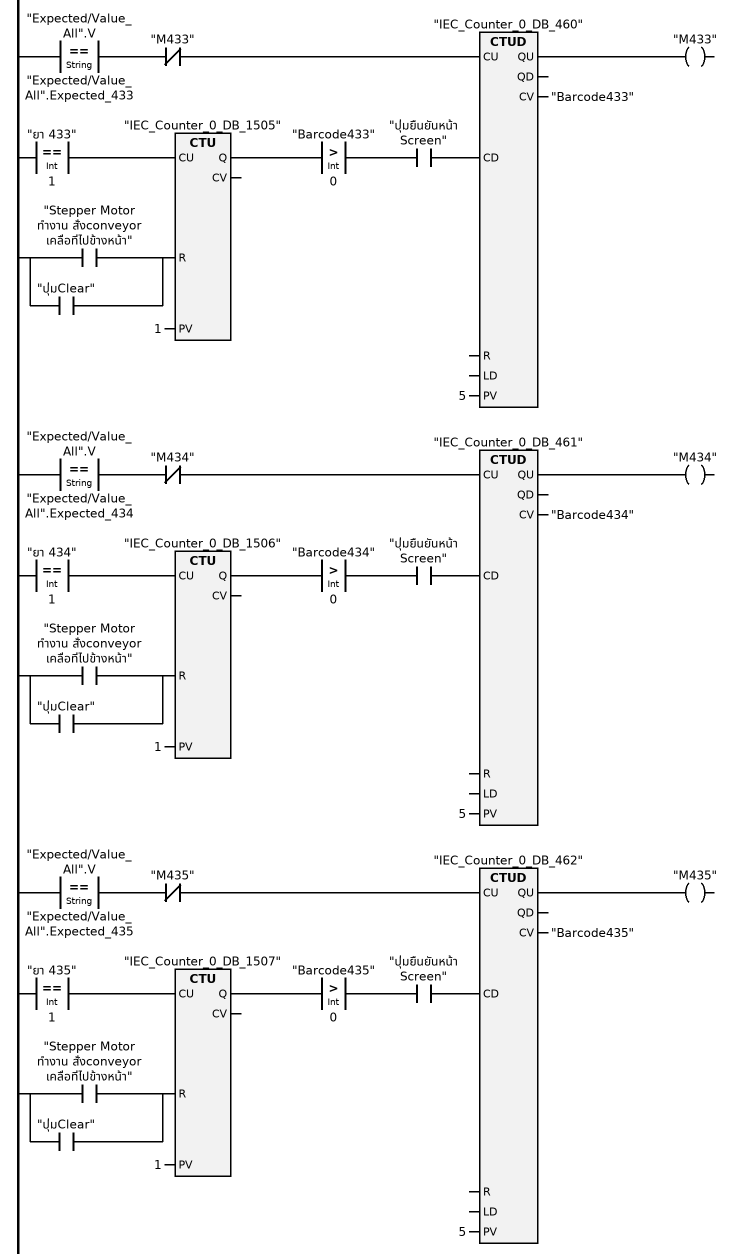
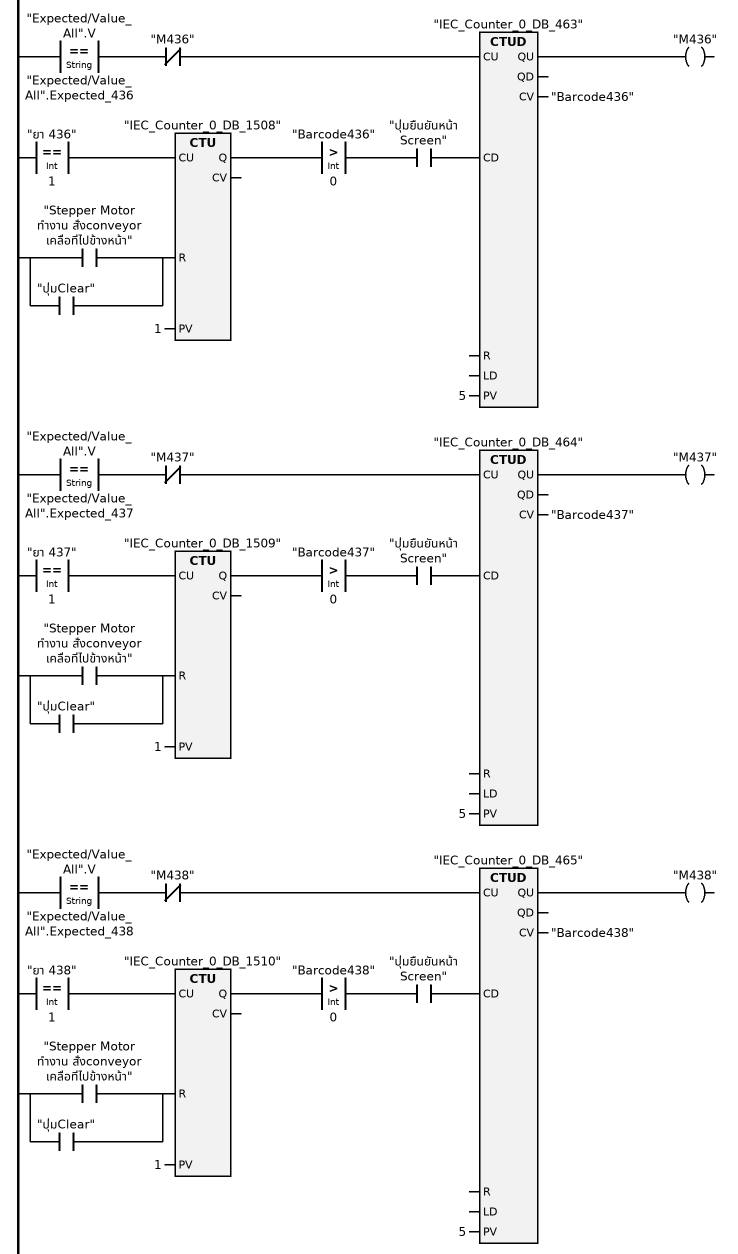
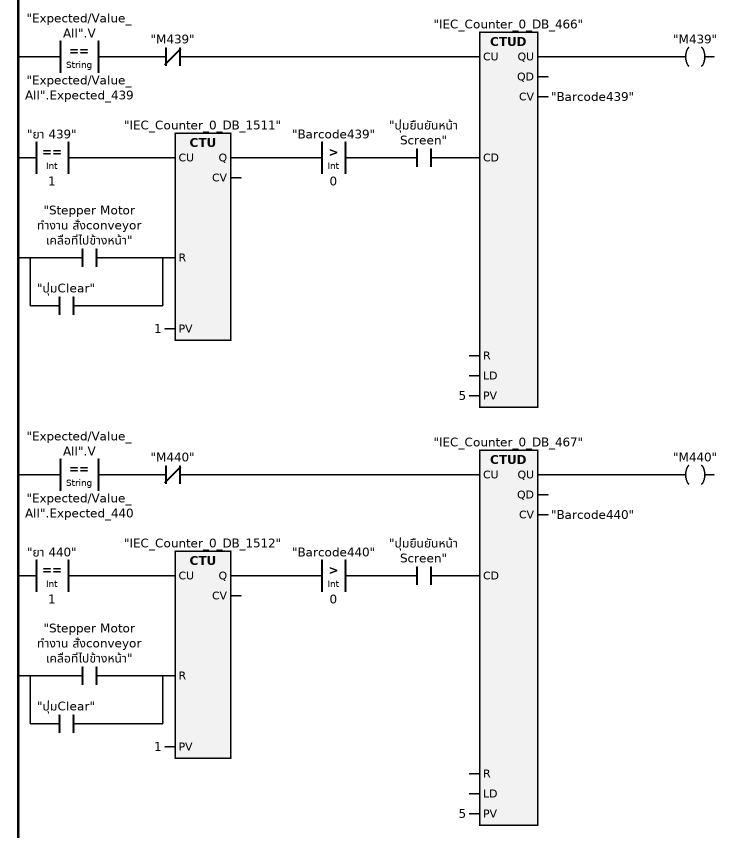
   "IEC_Counter_0_DB_1493".CTU(CU := "ยา 421" = 1,
                           R := "Stepper Motor ทำงาน สั่งconveyor เคลื่อที่ไปข้างหน้า" OR "ปุ่มClear",
                           PV := 1);
   "IEC_Counter_0_DB_448".CTUD(CU := ("Expected/Value_All".V = "Expected/Value_All".Expected_421) AND NOT "M421",
                           CD := "IEC_Counter_0_DB_1493".Q AND ("Barcode421" > 0) AND "ปุ่มยืนยันหน้า Screen",
                           PV := 5,
                           CV => "Barcode421");
   "M421" := "IEC_Counter_0_DB_448".QU;
   "IEC_Counter_0_DB_1494".CTU(CU := "ยา 422" = 1,
                           R := "Stepper Motor ทำงาน สั่งconveyor เคลื่อที่ไปข้างหน้า" OR "ปุ่มClear",
                           PV := 1);
   "IEC_Counter_0_DB_449".CTUD(CU := ("Expected/Value_All".V = "Expected/Value_All".Expected_422) AND NOT "M422",
                           CD := "IEC_Counter_0_DB_1494".Q AND ("Barcode422" > 0) AND "ปุ่มยืนยันหน้า Screen",
                           PV := 5,
                           CV => "Barcode422");
   "M422" := "IEC_Counter_0_DB_449".QU;
   "IEC_Counter_0_DB_1495".CTU(CU := "ยา 423" = 1,
                           R := "Stepper Motor ทำงาน สั่งconveyor เคลื่อที่ไปข้างหน้า" OR "ปุ่มClear",
                           PV := 1);
   "IEC_Counter_0_DB_450".CTUD(CU := ("Expected/Value_All".V = "Expected/Value_All".Expected_423) AND NOT "M423",
                           CD := "IEC_Counter_0_DB_1495".Q AND ("Barcode423" > 0) AND "ปุ่มยืนยันหน้า Screen",
                           PV := 5,
                           CV => "Barcode423");
   "M423" := "IEC_Counter_0_DB_450".QU;
   "IEC_Counter_0_DB_1496".CTU(CU := "ยา 424" = 1,
                           R := "Stepper Motor ทำงาน สั่งconveyor เคลื่อที่ไปข้างหน้า" OR "ปุ่มClear",
                           PV := 1);
   "IEC_Counter_0_DB_451".CTUD(CU := ("Expected/Value_All".V = "Expected/Value_All".Expected_424) AND NOT "M424",
                           CD := "IEC_Counter_0_DB_1496".Q AND ("Barcode424" > 0) AND "ปุ่มยืนยันหน้า Screen",
                           PV := 5,
                           CV => "Barcode424");
   "M424" := "IEC_Counter_0_DB_451".QU;
   "IEC_Counter_0_DB_1497".CTU(CU := "ยา 425" = 1,
                           R := "Stepper Motor ทำงาน สั่งconveyor เคลื่อที่ไปข้างหน้า" OR "ปุ่มClear",
                           PV := 1);
   "IEC_Counter_0_DB_452".CTUD(CU := ("Expected/Value_All".V = "Expected/Value_All".Expected_425) AND NOT "M425",
                           CD := "IEC_Counter_0_DB_1497".Q AND ("Barcode425" > 0) AND "ปุ่มยืนยันหน้า Screen",
                           PV := 5,
                           CV => "Barcode425");
   "M425" := "IEC_Counter_0_DB_452".QU;
   "IEC_Counter_0_DB_1498".CTU(CU := "ยา 426" = 1,
                           R := "Stepper Motor ทำงาน สั่งconveyor เคลื่อที่ไปข้างหน้า" OR "ปุ่มClear",
                           PV := 1);
   "IEC_Counter_0_DB_453".CTUD(CU := ("Expected/Value_All".V = "Expected/Value_All".Expected_426) AND NOT "M426",
                           CD := "IEC_Counter_0_DB_1498".Q AND ("Barcode426" > 0) AND "ปุ่มยืนยันหน้า Screen",
                           PV := 5,
                           CV => "Barcode426");
   "M426" := "IEC_Counter_0_DB_453".QU;
   "IEC_Counter_0_DB_1499".CTU(CU := "ยา 427" = 1,
                           R := "Stepper Motor ทำงาน สั่งconveyor เคลื่อที่ไปข้างหน้า" OR "ปุ่มClear",
                           PV := 1);
   "IEC_Counter_0_DB_454".CTUD(CU := ("Expected/Value_All".V = "Expected/Value_All".Expected_427) AND NOT "M427",
                           CD := "IEC_Counter_0_DB_1499".Q AND ("Barcode427" > 0) AND "ปุ่มยืนยันหน้า Screen",
                           PV := 5,
                           CV => "Barcode427");
   "M427" := "IEC_Counter_0_DB_454".QU;
   "IEC_Counter_0_DB_1500".CTU(CU := "ยา 428" = 1,
                           R := "Stepper Motor ทำงาน สั่งconveyor เคลื่อที่ไปข้างหน้า" OR "ปุ่มClear",
                           PV := 1);
   "IEC_Counter_0_DB_455".CTUD(CU := ("Expected/Value_All".V = "Expected/Value_All".Expected_428) AND NOT "M428",
                           CD := "IEC_Counter_0_DB_1500".Q AND ("Barcode428" > 0) AND "ปุ่มยืนยันหน้า Screen",
                           PV := 5,
                           CV => "Barcode428");
   "M428" := "IEC_Counter_0_DB_455".QU;
   "IEC_Counter_0_DB_1501".CTU(CU := "ยา 429" = 1,
                           R := "Stepper Motor ทำงาน สั่งconveyor เคลื่อที่ไปข้างหน้า" OR "ปุ่มClear",
                           PV := 1);
   "IEC_Counter_0_DB_456".CTUD(CU := ("Expected/Value_All".V = "Expected/Value_All".Expected_429) AND NOT "M429",
                           CD := "IEC_Counter_0_DB_1501".Q AND ("Barcode429" > 0) AND "ปุ่มยืนยันหน้า Screen",
                           PV := 5,
                           CV => "Barcode429");
   "M429" := "IEC_Counter_0_DB_456".QU;
   "IEC_Counter_0_DB_1502".CTU(CU := "ยา 430" = 1,
                           R := "Stepper Motor ทำงาน สั่งconveyor เคลื่อที่ไปข้างหน้า" OR "ปุ่มClear",
                           PV := 1);
   "IEC_Counter_0_DB_457".CTUD(CU := ("Expected/Value_All".V = "Expected/Value_All".Expected_430) AND NOT "M430",
                           CD := "IEC_Counter_0_DB_1502".Q AND ("Barcode430" > 0) AND "ปุ่มยืนยันหน้า Screen",
                           PV := 5,
                           CV => "Barcode430");
   "M430" := "IEC_Counter_0_DB_457".QU;
   "IEC_Counter_0_DB_1503".CTU(CU := "ยา 431" = 1,
                           R := "Stepper Motor ทำงาน สั่งconveyor เคลื่อที่ไปข้างหน้า" OR "ปุ่มClear",
                           PV := 1);
   "IEC_Counter_0_DB_458".CTUD(CU := ("Expected/Value_All".V = "Expected/Value_All".Expected_431) AND NOT "M431",
                           CD := "IEC_Counter_0_DB_1503".Q AND ("Barcode431" > 0) AND "ปุ่มยืนยันหน้า Screen",
                           PV := 5,
                           CV => "Barcode431");
   "M431" := "IEC_Counter_0_DB_458".QU;
   "IEC_Counter_0_DB_1504".CTU(CU := "ยา 432" = 1,
                           R := "Stepper Motor ทำงาน สั่งconveyor เคลื่อที่ไปข้างหน้า" OR "ปุ่มClear",
                           PV := 1);
   "IEC_Counter_0_DB_459".CTUD(CU := ("Expected/Value_All".V = "Expected/Value_All".Expected_432) AND NOT "M432",
                           CD := "IEC_Counter_0_DB_1504".Q AND ("Barcode432" > 0) AND "ปุ่มยืนยันหน้า Screen",
                           PV := 5,
                           CV => "Barcode432");
   "M432" := "IEC_Counter_0_DB_459".QU;
   "IEC_Counter_0_DB_1505".CTU(CU := "ยา 433" = 1,
                           R := "Stepper Motor ทำงาน สั่งconveyor เคลื่อที่ไปข้างหน้า" OR "ปุ่มClear",
                           PV := 1);
   "IEC_Counter_0_DB_460".CTUD(CU := ("Expected/Value_All".V = "Expected/Value_All".Expected_433) AND NOT "M433",
                           CD := "IEC_Counter_0_DB_1505".Q AND ("Barcode433" > 0) AND "ปุ่มยืนยันหน้า Screen",
                           PV := 5,
                           CV => "Barcode433");
   "M433" := "IEC_Counter_0_DB_460".QU;
   "IEC_Counter_0_DB_1506".CTU(CU := "ยา 434" = 1,
                           R := "Stepper Motor ทำงาน สั่งconveyor เคลื่อที่ไปข้างหน้า" OR "ปุ่มClear",
                           PV := 1);
   "IEC_Counter_0_DB_461".CTUD(CU := ("Expected/Value_All".V = "Expected/Value_All".Expected_434) AND NOT "M434",
                           CD := "IEC_Counter_0_DB_1506".Q AND ("Barcode434" > 0) AND "ปุ่มยืนยันหน้า Screen",
                           PV := 5,
                           CV => "Barcode434");
   "M434" := "IEC_Counter_0_DB_461".QU;
   "IEC_Counter_0_DB_1507".CTU(CU := "ยา 435" = 1,
                           R := "Stepper Motor ทำงาน สั่งconveyor เคลื่อที่ไปข้างหน้า" OR "ปุ่มClear",
                           PV := 1);
   "IEC_Counter_0_DB_462".CTUD(CU := ("Expected/Value_All".V = "Expected/Value_All".Expected_435) AND NOT "M435",
                           CD := "IEC_Counter_0_DB_1507".Q AND ("Barcode435" > 0) AND "ปุ่มยืนยันหน้า Screen",
                           PV := 5,
                           CV => "Barcode435");
   "M435" := "IEC_Counter_0_DB_462".QU;
   "IEC_Counter_0_DB_1508".CTU(CU := "ยา 436" = 1,
                           R := "Stepper Motor ทำงาน สั่งconveyor เคลื่อที่ไปข้างหน้า" OR "ปุ่มClear",
                           PV := 1);
   "IEC_Counter_0_DB_463".CTUD(CU := ("Expected/Value_All".V = "Expected/Value_All".Expected_436) AND NOT "M436",
                           CD := "IEC_Counter_0_DB_1508".Q AND ("Barcode436" > 0) AND "ปุ่มยืนยันหน้า Screen",
                           PV := 5,
                           CV => "Barcode436");
   "M436" := "IEC_Counter_0_DB_463".QU;
   "IEC_Counter_0_DB_1509".CTU(CU := "ยา 437" = 1,
                           R := "Stepper Motor ทำงาน สั่งconveyor เคลื่อที่ไปข้างหน้า" OR "ปุ่มClear",
                           PV := 1);
   "IEC_Counter_0_DB_464".CTUD(CU := ("Expected/Value_All".V = "Expected/Value_All".Expected_437) AND NOT "M437",
                           CD := "IEC_Counter_0_DB_1509".Q AND ("Barcode437" > 0) AND "ปุ่มยืนยันหน้า Screen",
                           PV := 5,
                           CV => "Barcode437");
   "M437" := "IEC_Counter_0_DB_464".QU;
   "IEC_Counter_0_DB_1510".CTU(CU := "ยา 438" = 1,
                           R := "Stepper Motor ทำงาน สั่งconveyor เคลื่อที่ไปข้างหน้า" OR "ปุ่มClear",
                           PV := 1);
   "IEC_Counter_0_DB_465".CTUD(CU := ("Expected/Value_All".V = "Expected/Value_All".Expected_438) AND NOT "M438",
                           CD := "IEC_Counter_0_DB_1510".Q AND ("Barcode438" > 0) AND "ปุ่มยืนยันหน้า Screen",
                           PV := 5,
                           CV => "Barcode438");
   "M438" := "IEC_Counter_0_DB_465".QU;
   "IEC_Counter_0_DB_1511".CTU(CU := "ยา 439" = 1,
                           R := "Stepper Motor ทำงาน สั่งconveyor เคลื่อที่ไปข้างหน้า" OR "ปุ่มClear",
                           PV := 1);
   "IEC_Counter_0_DB_466".CTUD(CU := ("Expected/Value_All".V = "Expected/Value_All".Expected_439) AND NOT "M439",
                           CD := "IEC_Counter_0_DB_1511".Q AND ("Barcode439" > 0) AND "ปุ่มยืนยันหน้า Screen",
                           PV := 5,
                           CV => "Barcode439");
   "M439" := "IEC_Counter_0_DB_466".QU;
   "IEC_Counter_0_DB_1512".CTU(CU := "ยา 440" = 1,
                           R := "Stepper Motor ทำงาน สั่งconveyor เคลื่อที่ไปข้างหน้า" OR "ปุ่มClear",
                           PV := 1);
   "IEC_Counter_0_DB_467".CTUD(CU := ("Expected/Value_All".V = "Expected/Value_All".Expected_440) AND NOT "M440",
                           CD := "IEC_Counter_0_DB_1512".Q AND ("Barcode440" > 0) AND "ปุ่มยืนยันหน้า Screen",
                           PV := 5,
                           CV => "Barcode440");
   "M440" := "IEC_Counter_0_DB_467".QU;
END_REGION

REGION Network 23
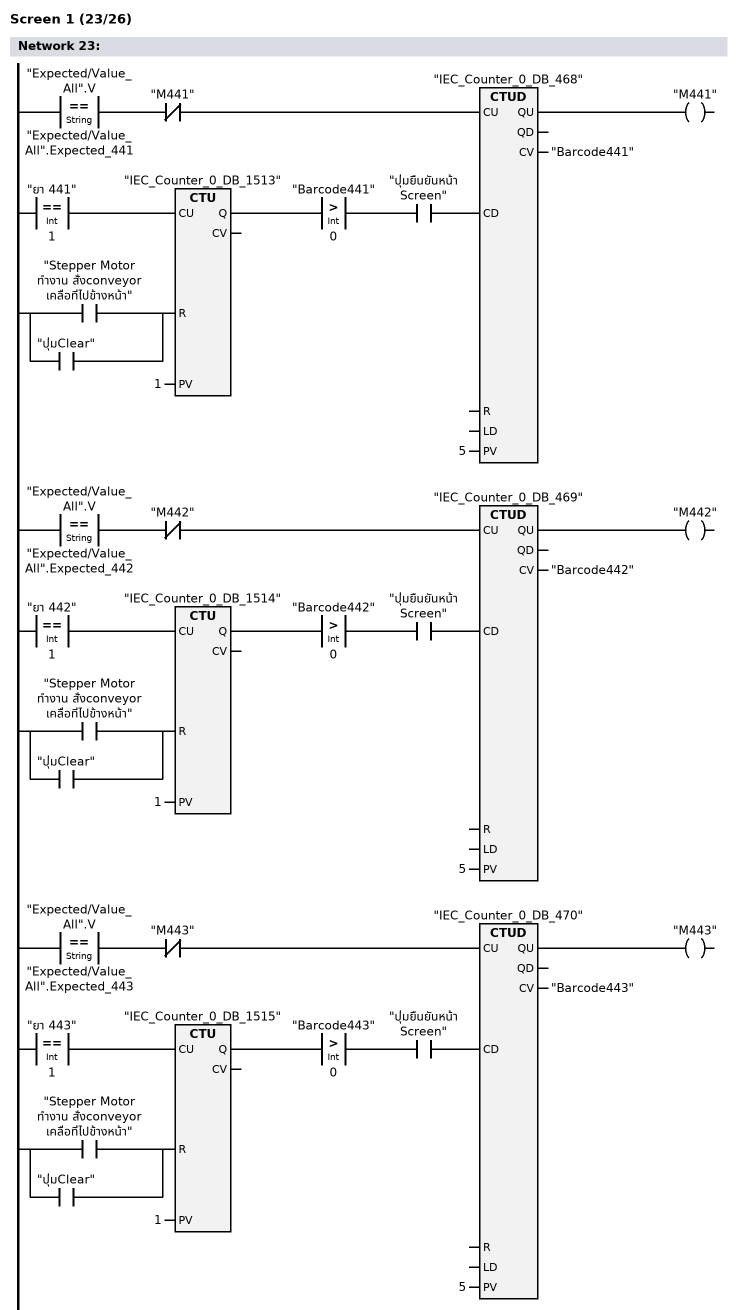
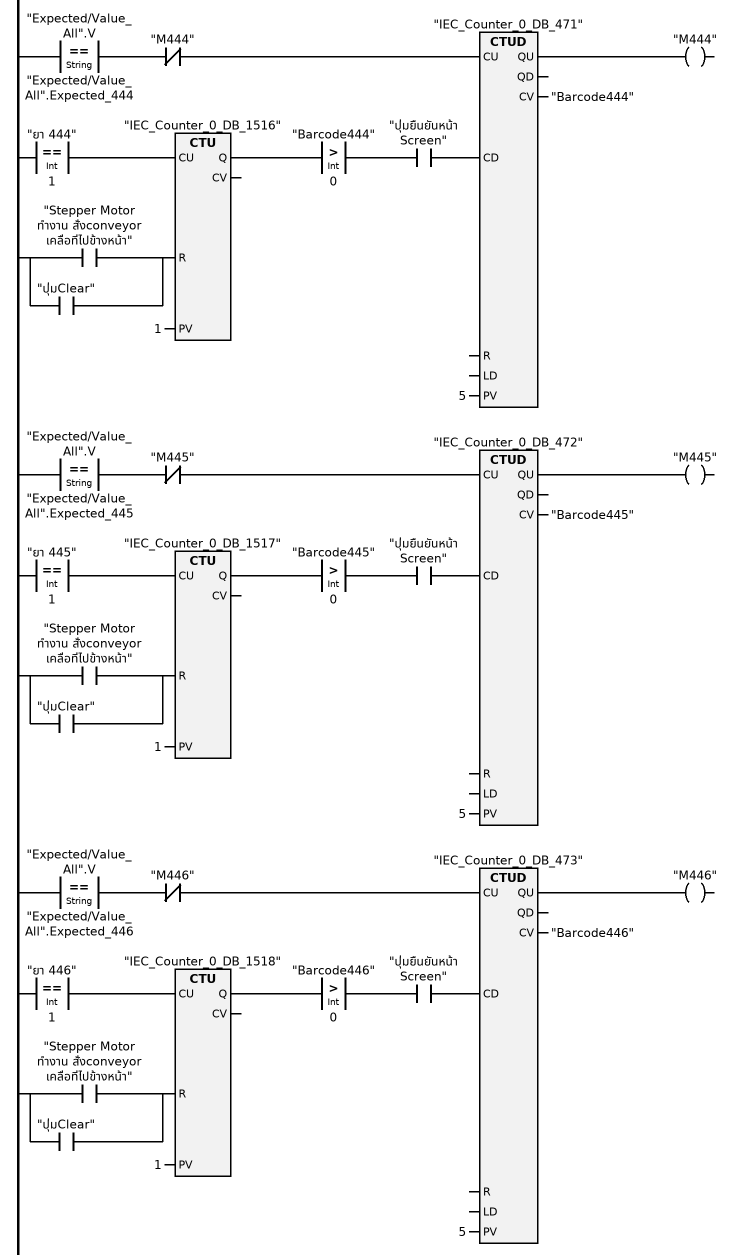
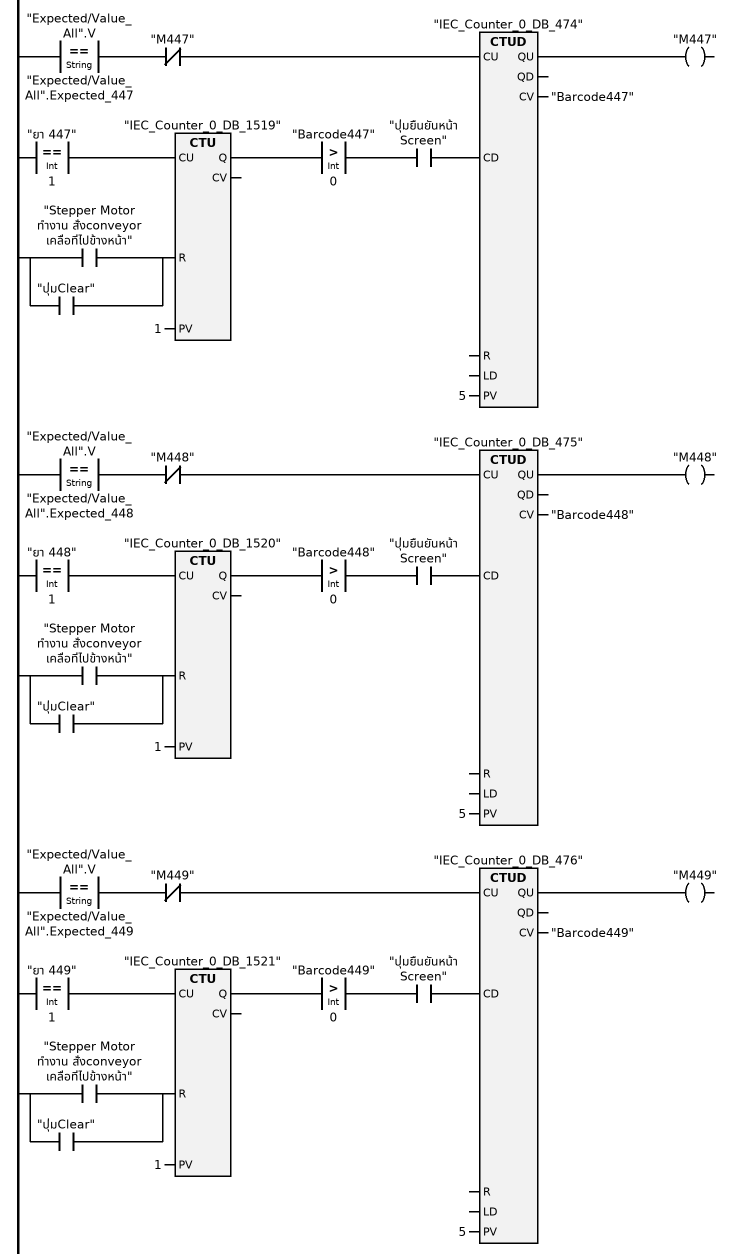
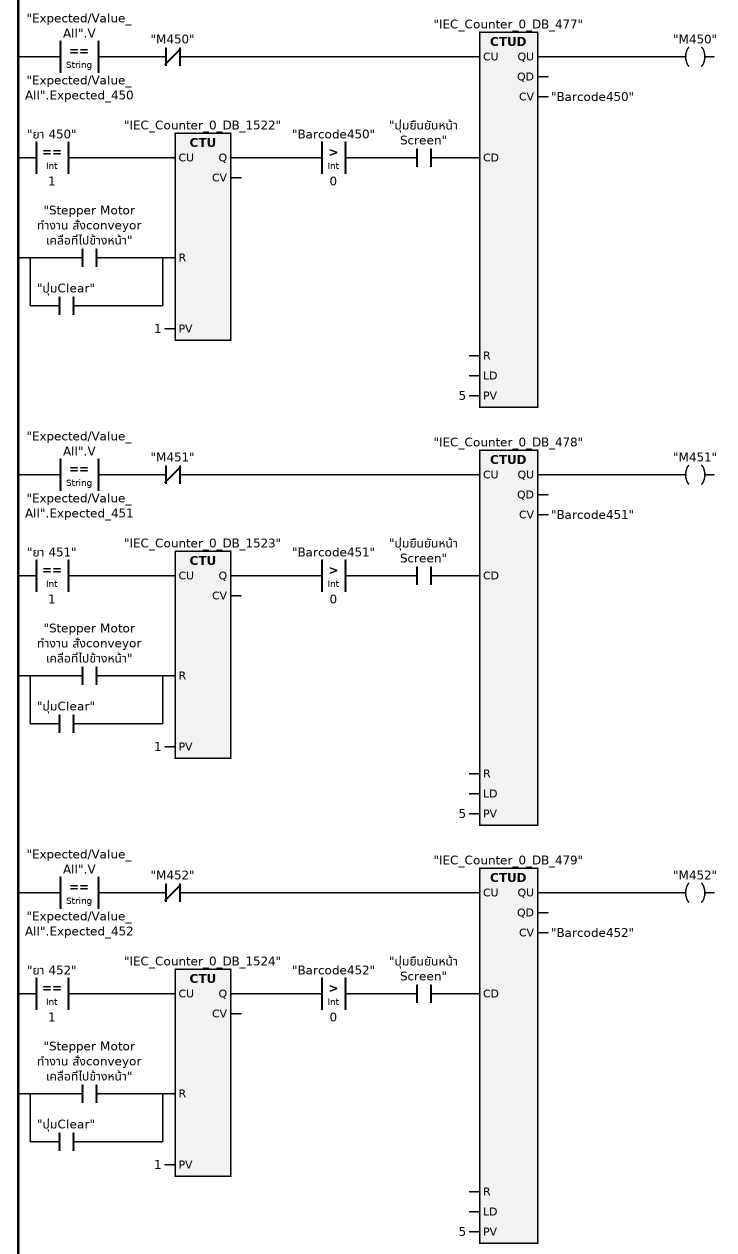
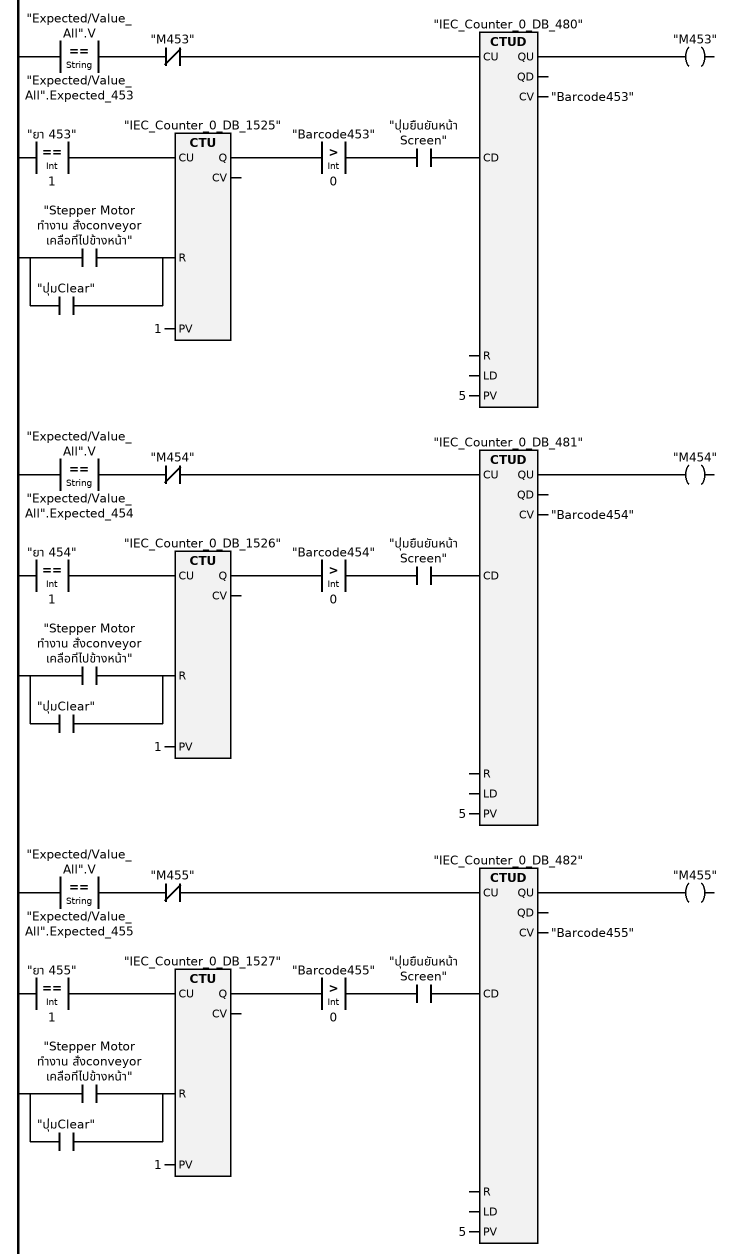
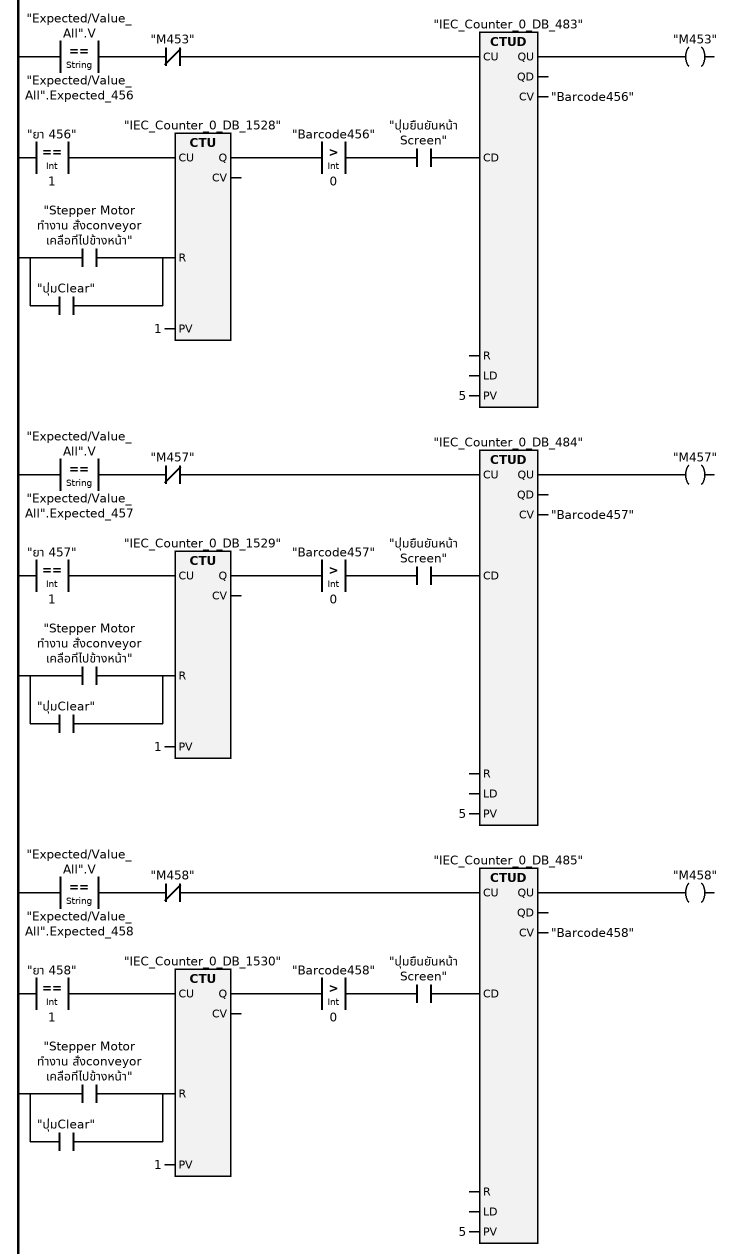
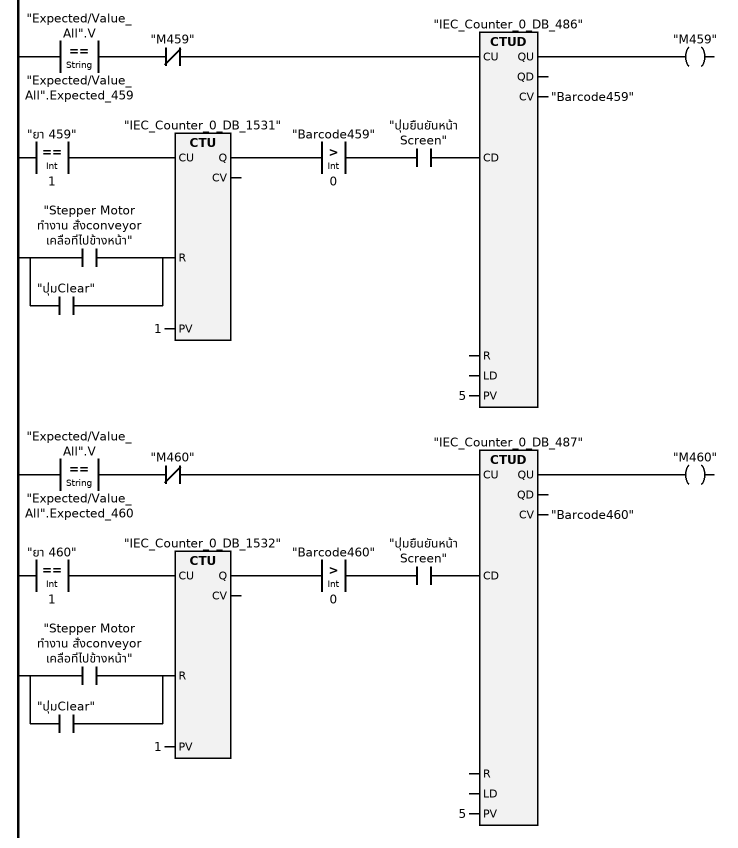
   "IEC_Counter_0_DB_1513".CTU(CU := "ยา 441" = 1,
                           R := "Stepper Motor ทำงาน สั่งconveyor เคลื่อที่ไปข้างหน้า" OR "ปุ่มClear",
                           PV := 1);
   "IEC_Counter_0_DB_468".CTUD(CU := ("Expected/Value_All".V = "Expected/Value_All".Expected_441) AND NOT "M441",
                           CD := "IEC_Counter_0_DB_1513".Q AND ("Barcode441" > 0) AND "ปุ่มยืนยันหน้า Screen",
                           PV := 5,
                           CV => "Barcode441");
   "M441" := "IEC_Counter_0_DB_468".QU;
   "IEC_Counter_0_DB_1514".CTU(CU := "ยา 442" = 1,
                           R := "Stepper Motor ทำงาน สั่งconveyor เคลื่อที่ไปข้างหน้า" OR "ปุ่มClear",
                           PV := 1);
   "IEC_Counter_0_DB_469".CTUD(CU := ("Expected/Value_All".V = "Expected/Value_All".Expected_442) AND NOT "M442",
                           CD := "IEC_Counter_0_DB_1514".Q AND ("Barcode442" > 0) AND "ปุ่มยืนยันหน้า Screen",
                           PV := 5,
                           CV => "Barcode442");
   "M442" := "IEC_Counter_0_DB_469".QU;
   "IEC_Counter_0_DB_1515".CTU(CU := "ยา 443" = 1,
                           R := "Stepper Motor ทำงาน สั่งconveyor เคลื่อที่ไปข้างหน้า" OR "ปุ่มClear",
                           PV := 1);
   "IEC_Counter_0_DB_470".CTUD(CU := ("Expected/Value_All".V = "Expected/Value_All".Expected_443) AND NOT "M443",
                           CD := "IEC_Counter_0_DB_1515".Q AND ("Barcode443" > 0) AND "ปุ่มยืนยันหน้า Screen",
                           PV := 5,
                           CV => "Barcode443");
   "M443" := "IEC_Counter_0_DB_470".QU;
   "IEC_Counter_0_DB_1516".CTU(CU := "ยา 444" = 1,
                           R := "Stepper Motor ทำงาน สั่งconveyor เคลื่อที่ไปข้างหน้า" OR "ปุ่มClear",
                           PV := 1);
   "IEC_Counter_0_DB_471".CTUD(CU := ("Expected/Value_All".V = "Expected/Value_All".Expected_444) AND NOT "M444",
                           CD := "IEC_Counter_0_DB_1516".Q AND ("Barcode444" > 0) AND "ปุ่มยืนยันหน้า Screen",
                           PV := 5,
                           CV => "Barcode444");
   "M444" := "IEC_Counter_0_DB_471".QU;
   "IEC_Counter_0_DB_1517".CTU(CU := "ยา 445" = 1,
                           R := "Stepper Motor ทำงาน สั่งconveyor เคลื่อที่ไปข้างหน้า" OR "ปุ่มClear",
                           PV := 1);
   "IEC_Counter_0_DB_472".CTUD(CU := ("Expected/Value_All".V = "Expected/Value_All".Expected_445) AND NOT "M445",
                           CD := "IEC_Counter_0_DB_1517".Q AND ("Barcode445" > 0) AND "ปุ่มยืนยันหน้า Screen",
                           PV := 5,
                           CV => "Barcode445");
   "M445" := "IEC_Counter_0_DB_472".QU;
   "IEC_Counter_0_DB_1518".CTU(CU := "ยา 446" = 1,
                           R := "Stepper Motor ทำงาน สั่งconveyor เคลื่อที่ไปข้างหน้า" OR "ปุ่มClear",
                           PV := 1);
   "IEC_Counter_0_DB_473".CTUD(CU := ("Expected/Value_All".V = "Expected/Value_All".Expected_446) AND NOT "M446",
                           CD := "IEC_Counter_0_DB_1518".Q AND ("Barcode446" > 0) AND "ปุ่มยืนยันหน้า Screen",
                           PV := 5,
                           CV => "Barcode446");
   "M446" := "IEC_Counter_0_DB_473".QU;
   "IEC_Counter_0_DB_1519".CTU(CU := "ยา 447" = 1,
                           R := "Stepper Motor ทำงาน สั่งconveyor เคลื่อที่ไปข้างหน้า" OR "ปุ่มClear",
                           PV := 1);
   "IEC_Counter_0_DB_474".CTUD(CU := ("Expected/Value_All".V = "Expected/Value_All".Expected_447) AND NOT "M447",
                           CD := "IEC_Counter_0_DB_1519".Q AND ("Barcode447" > 0) AND "ปุ่มยืนยันหน้า Screen",
                           PV := 5,
                           CV => "Barcode447");
   "M447" := "IEC_Counter_0_DB_474".QU;
   "IEC_Counter_0_DB_1520".CTU(CU := "ยา 448" = 1,
                           R := "Stepper Motor ทำงาน สั่งconveyor เคลื่อที่ไปข้างหน้า" OR "ปุ่มClear",
                           PV := 1);
   "IEC_Counter_0_DB_475".CTUD(CU := ("Expected/Value_All".V = "Expected/Value_All".Expected_448) AND NOT "M448",
                           CD := "IEC_Counter_0_DB_1520".Q AND ("Barcode448" > 0) AND "ปุ่มยืนยันหน้า Screen",
                           PV := 5,
                           CV => "Barcode448");
   "M448" := "IEC_Counter_0_DB_475".QU;
   "IEC_Counter_0_DB_1521".CTU(CU := "ยา 449" = 1,
                           R := "Stepper Motor ทำงาน สั่งconveyor เคลื่อที่ไปข้างหน้า" OR "ปุ่มClear",
                           PV := 1);
   "IEC_Counter_0_DB_476".CTUD(CU := ("Expected/Value_All".V = "Expected/Value_All".Expected_449) AND NOT "M449",
                           CD := "IEC_Counter_0_DB_1521".Q AND ("Barcode449" > 0) AND "ปุ่มยืนยันหน้า Screen",
                           PV := 5,
                           CV => "Barcode449");
   "M449" := "IEC_Counter_0_DB_476".QU;
   "IEC_Counter_0_DB_1522".CTU(CU := "ยา 450" = 1,
                           R := "Stepper Motor ทำงาน สั่งconveyor เคลื่อที่ไปข้างหน้า" OR "ปุ่มClear",
                           PV := 1);
   "IEC_Counter_0_DB_477".CTUD(CU := ("Expected/Value_All".V = "Expected/Value_All".Expected_450) AND NOT "M450",
                           CD := "IEC_Counter_0_DB_1522".Q AND ("Barcode450" > 0) AND "ปุ่มยืนยันหน้า Screen",
                           PV := 5,
                           CV => "Barcode450");
   "M450" := "IEC_Counter_0_DB_477".QU;
   "IEC_Counter_0_DB_1523".CTU(CU := "ยา 451" = 1,
                           R := "Stepper Motor ทำงาน สั่งconveyor เคลื่อที่ไปข้างหน้า" OR "ปุ่มClear",
                           PV := 1);
   "IEC_Counter_0_DB_478".CTUD(CU := ("Expected/Value_All".V = "Expected/Value_All".Expected_451) AND NOT "M451",
                           CD := "IEC_Counter_0_DB_1523".Q AND ("Barcode451" > 0) AND "ปุ่มยืนยันหน้า Screen",
                           PV := 5,
                           CV => "Barcode451");
   "M451" := "IEC_Counter_0_DB_478".QU;
   "IEC_Counter_0_DB_1524".CTU(CU := "ยา 452" = 1,
                           R := "Stepper Motor ทำงาน สั่งconveyor เคลื่อที่ไปข้างหน้า" OR "ปุ่มClear",
                           PV := 1);
   "IEC_Counter_0_DB_479".CTUD(CU := ("Expected/Value_All".V = "Expected/Value_All".Expected_452) AND NOT "M452",
                           CD := "IEC_Counter_0_DB_1524".Q AND ("Barcode452" > 0) AND "ปุ่มยืนยันหน้า Screen",
                           PV := 5,
                           CV => "Barcode452");
   "M452" := "IEC_Counter_0_DB_479".QU;
   "IEC_Counter_0_DB_1525".CTU(CU := "ยา 453" = 1,
                           R := "Stepper Motor ทำงาน สั่งconveyor เคลื่อที่ไปข้างหน้า" OR "ปุ่มClear",
                           PV := 1);
   "IEC_Counter_0_DB_480".CTUD(CU := ("Expected/Value_All".V = "Expected/Value_All".Expected_453) AND NOT "M453",
                           CD := "IEC_Counter_0_DB_1525".Q AND ("Barcode453" > 0) AND "ปุ่มยืนยันหน้า Screen",
                           PV := 5,
                           CV => "Barcode453");
   "M453" := "IEC_Counter_0_DB_480".QU;
   "IEC_Counter_0_DB_1526".CTU(CU := "ยา 454" = 1,
                           R := "Stepper Motor ทำงาน สั่งconveyor เคลื่อที่ไปข้างหน้า" OR "ปุ่มClear",
                           PV := 1);
   "IEC_Counter_0_DB_481".CTUD(CU := ("Expected/Value_All".V = "Expected/Value_All".Expected_454) AND NOT "M454",
                           CD := "IEC_Counter_0_DB_1526".Q AND ("Barcode454" > 0) AND "ปุ่มยืนยันหน้า Screen",
                           PV := 5,
                           CV => "Barcode454");
   "M454" := "IEC_Counter_0_DB_481".QU;
   "IEC_Counter_0_DB_1527".CTU(CU := "ยา 455" = 1,
                           R := "Stepper Motor ทำงาน สั่งconveyor เคลื่อที่ไปข้างหน้า" OR "ปุ่มClear",
                           PV := 1);
   "IEC_Counter_0_DB_482".CTUD(CU := ("Expected/Value_All".V = "Expected/Value_All".Expected_455) AND NOT "M455",
                           CD := "IEC_Counter_0_DB_1527".Q AND ("Barcode455" > 0) AND "ปุ่มยืนยันหน้า Screen",
                           PV := 5,
                           CV => "Barcode455");
   "M455" := "IEC_Counter_0_DB_482".QU;
   "IEC_Counter_0_DB_1528".CTU(CU := "ยา 456" = 1,
                           R := "Stepper Motor ทำงาน สั่งconveyor เคลื่อที่ไปข้างหน้า" OR "ปุ่มClear",
                           PV := 1);
   "IEC_Counter_0_DB_483".CTUD(CU := ("Expected/Value_All".V = "Expected/Value_All".Expected_456) AND NOT "M453",
                           CD := "IEC_Counter_0_DB_1528".Q AND ("Barcode456" > 0) AND "ปุ่มยืนยันหน้า Screen",
                           PV := 5,
                           CV => "Barcode456");
   "M453" := "IEC_Counter_0_DB_483".QU;
   "IEC_Counter_0_DB_1529".CTU(CU := "ยา 457" = 1,
                           R := "Stepper Motor ทำงาน สั่งconveyor เคลื่อที่ไปข้างหน้า" OR "ปุ่มClear",
                           PV := 1);
   "IEC_Counter_0_DB_484".CTUD(CU := ("Expected/Value_All".V = "Expected/Value_All".Expected_457) AND NOT "M457",
                           CD := "IEC_Counter_0_DB_1529".Q AND ("Barcode457" > 0) AND "ปุ่มยืนยันหน้า Screen",
                           PV := 5,
                           CV => "Barcode457");
   "M457" := "IEC_Counter_0_DB_484".QU;
   "IEC_Counter_0_DB_1530".CTU(CU := "ยา 458" = 1,
                           R := "Stepper Motor ทำงาน สั่งconveyor เคลื่อที่ไปข้างหน้า" OR "ปุ่มClear",
                           PV := 1);
   "IEC_Counter_0_DB_485".CTUD(CU := ("Expected/Value_All".V = "Expected/Value_All".Expected_458) AND NOT "M458",
                           CD := "IEC_Counter_0_DB_1530".Q AND ("Barcode458" > 0) AND "ปุ่มยืนยันหน้า Screen",
                           PV := 5,
                           CV => "Barcode458");
   "M458" := "IEC_Counter_0_DB_485".QU;
   "IEC_Counter_0_DB_1531".CTU(CU := "ยา 459" = 1,
                           R := "Stepper Motor ทำงาน สั่งconveyor เคลื่อที่ไปข้างหน้า" OR "ปุ่มClear",
                           PV := 1);
   "IEC_Counter_0_DB_486".CTUD(CU := ("Expected/Value_All".V = "Expected/Value_All".Expected_459) AND NOT "M459",
                           CD := "IEC_Counter_0_DB_1531".Q AND ("Barcode459" > 0) AND "ปุ่มยืนยันหน้า Screen",
                           PV := 5,
                           CV => "Barcode459");
   "M459" := "IEC_Counter_0_DB_486".QU;
   "IEC_Counter_0_DB_1532".CTU(CU := "ยา 460" = 1,
                           R := "Stepper Motor ทำงาน สั่งconveyor เคลื่อที่ไปข้างหน้า" OR "ปุ่มClear",
                           PV := 1);
   "IEC_Counter_0_DB_487".CTUD(CU := ("Expected/Value_All".V = "Expected/Value_All".Expected_460) AND NOT "M460",
                           CD := "IEC_Counter_0_DB_1532".Q AND ("Barcode460" > 0) AND "ปุ่มยืนยันหน้า Screen",
                           PV := 5,
                           CV => "Barcode460");
   "M460" := "IEC_Counter_0_DB_487".QU;
END_REGION

REGION Network 24
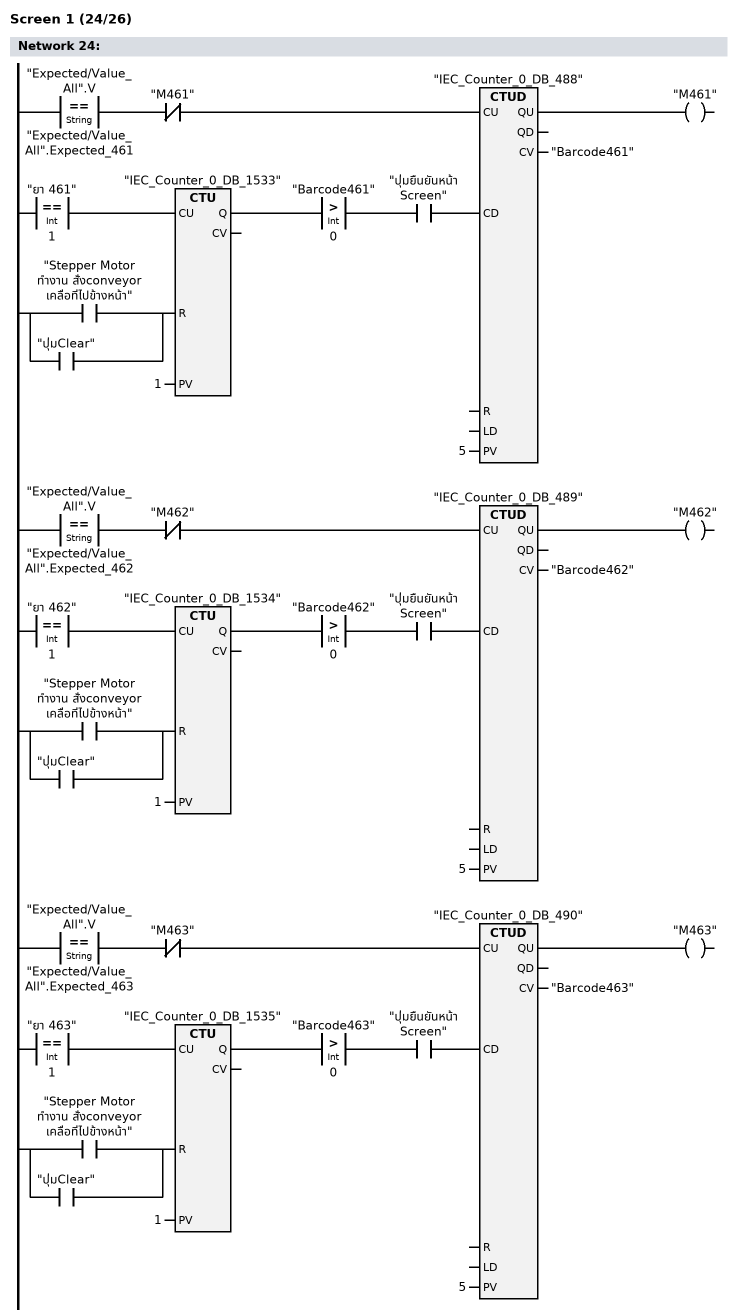
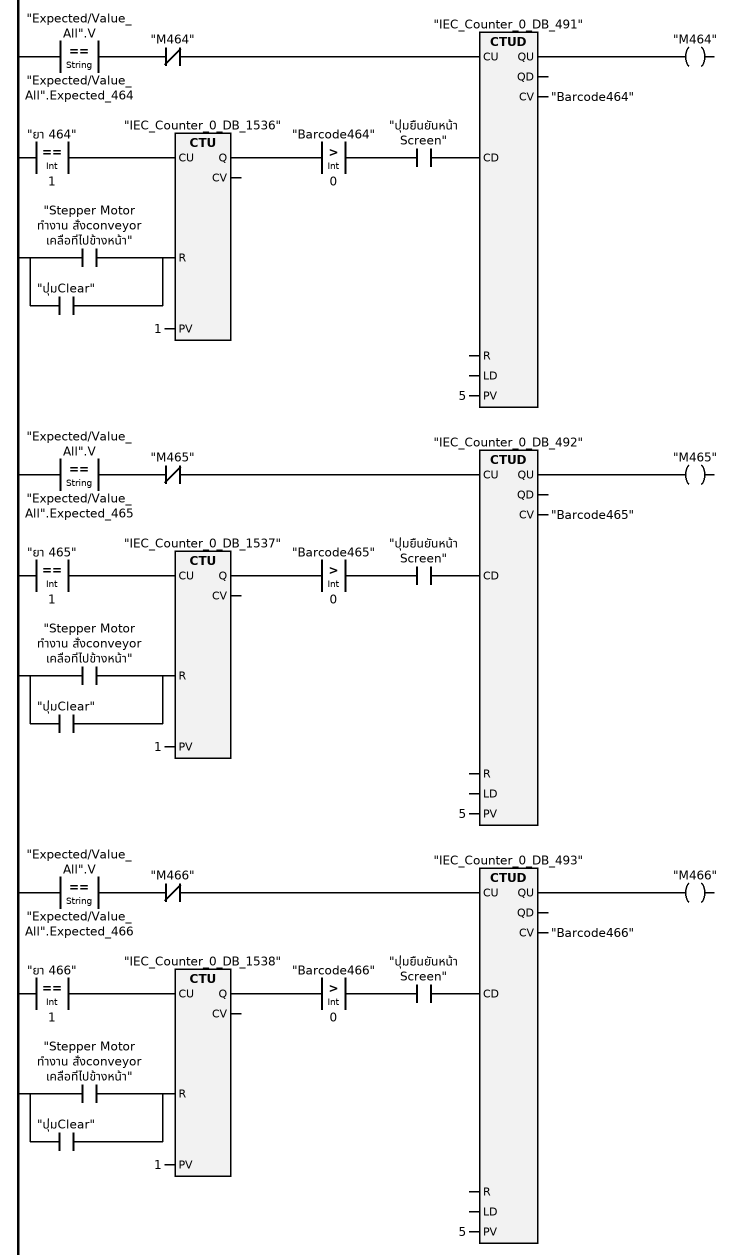
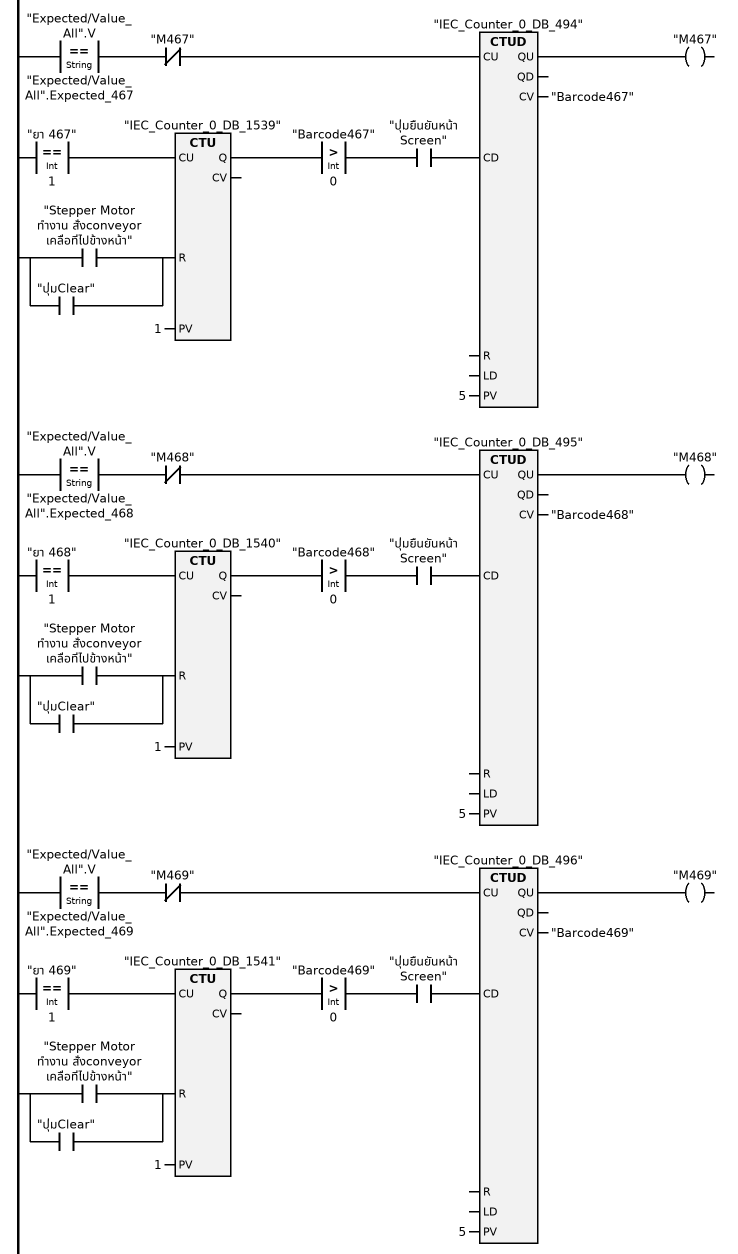
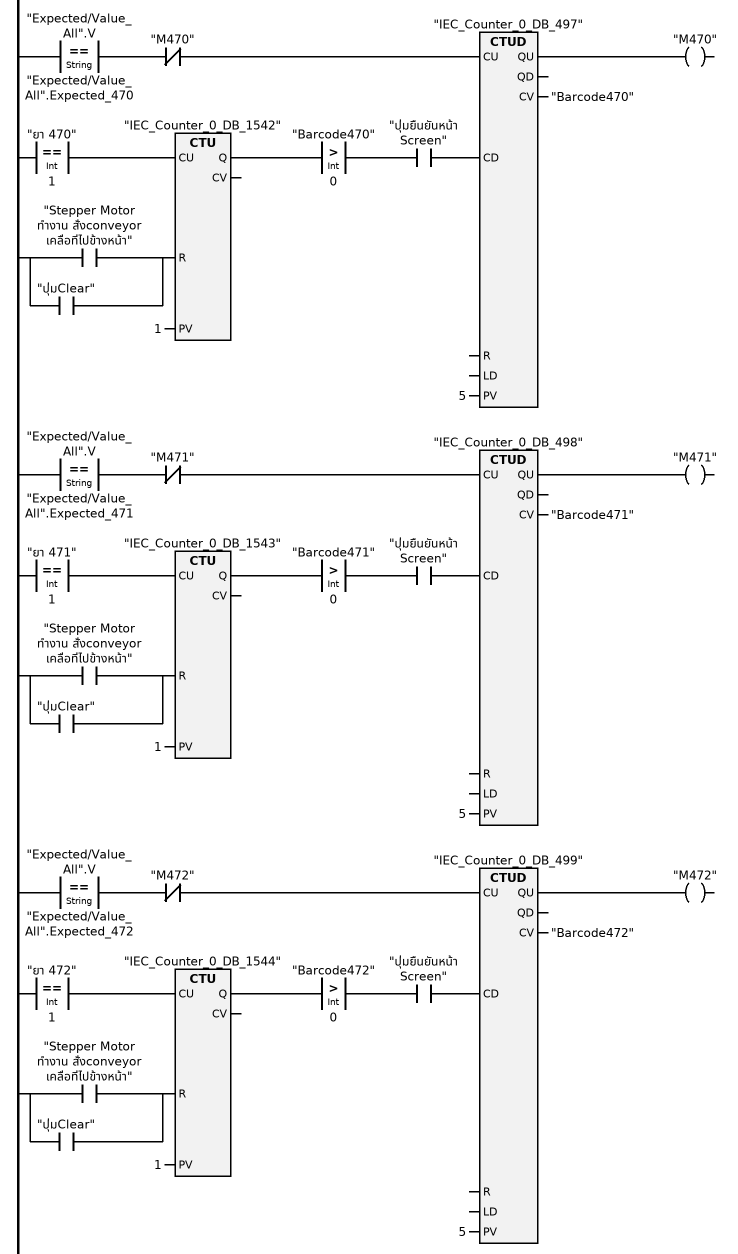
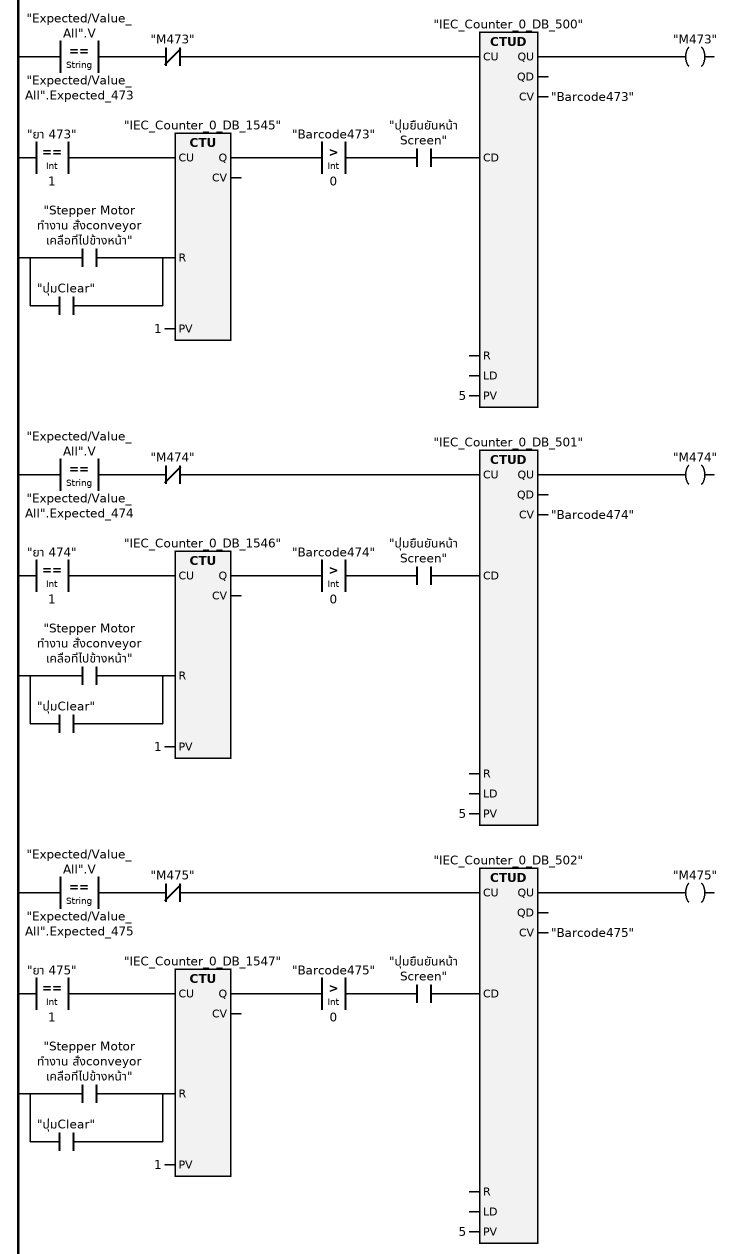
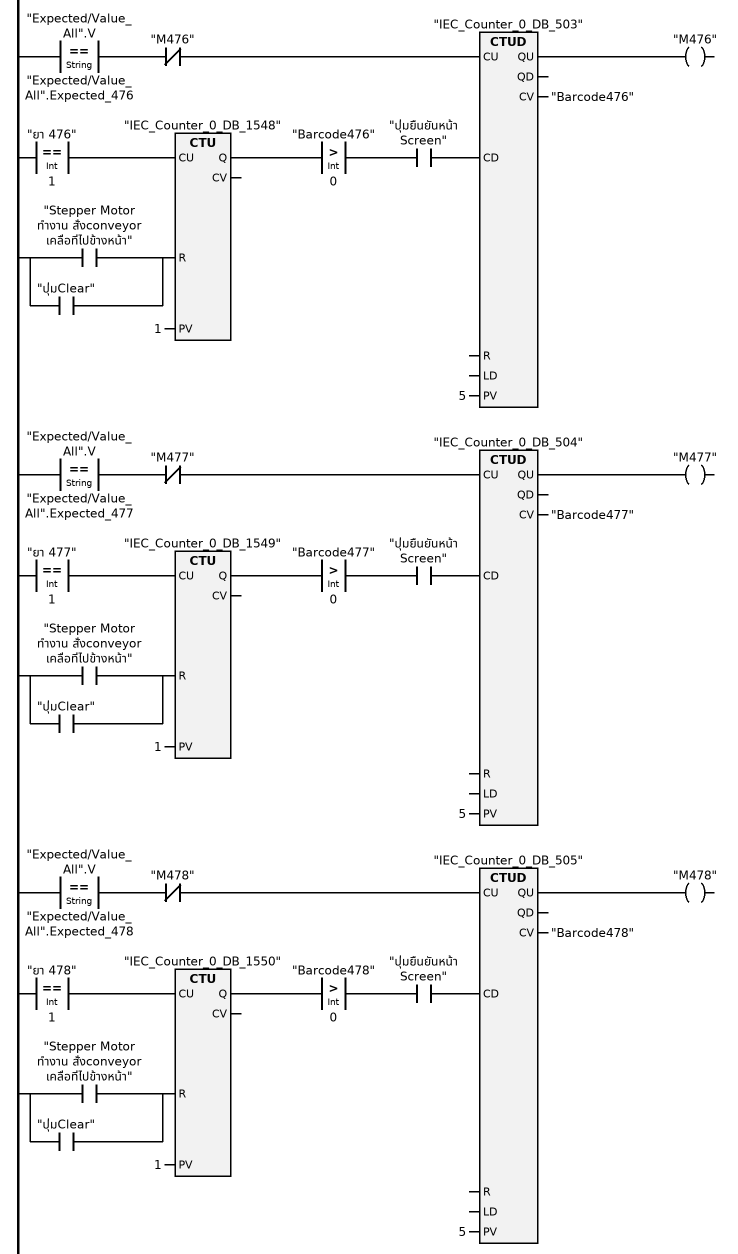
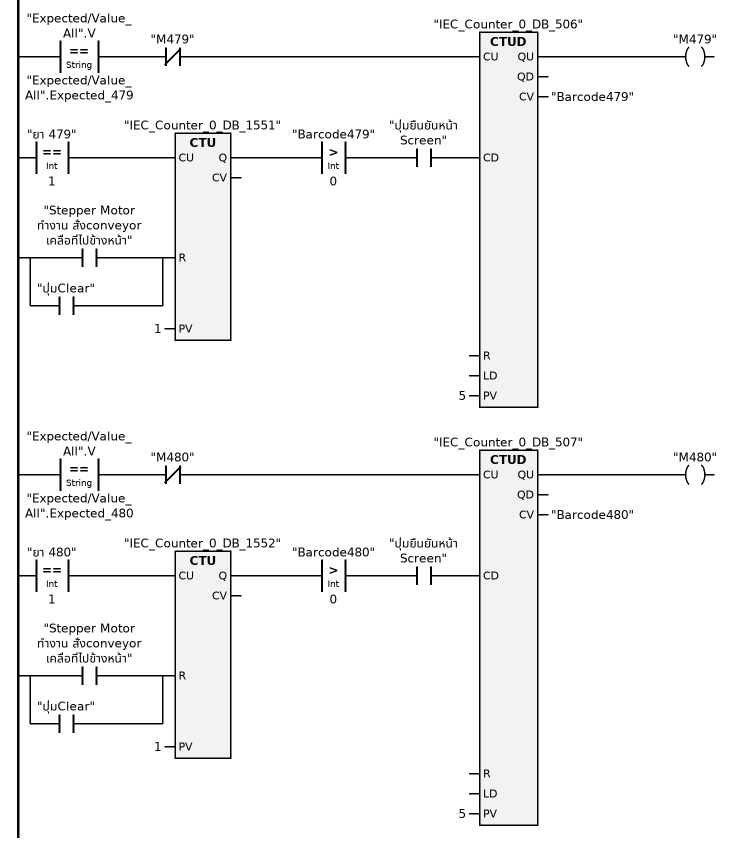
   "IEC_Counter_0_DB_1533".CTU(CU := "ยา 461" = 1,
                           R := "Stepper Motor ทำงาน สั่งconveyor เคลื่อที่ไปข้างหน้า" OR "ปุ่มClear",
                           PV := 1);
   "IEC_Counter_0_DB_488".CTUD(CU := ("Expected/Value_All".V = "Expected/Value_All".Expected_461) AND NOT "M461",
                           CD := "IEC_Counter_0_DB_1533".Q AND ("Barcode461" > 0) AND "ปุ่มยืนยันหน้า Screen",
                           PV := 5,
                           CV => "Barcode461");
   "M461" := "IEC_Counter_0_DB_488".QU;
   "IEC_Counter_0_DB_1534".CTU(CU := "ยา 462" = 1,
                           R := "Stepper Motor ทำงาน สั่งconveyor เคลื่อที่ไปข้างหน้า" OR "ปุ่มClear",
                           PV := 1);
   "IEC_Counter_0_DB_489".CTUD(CU := ("Expected/Value_All".V = "Expected/Value_All".Expected_462) AND NOT "M462",
                           CD := "IEC_Counter_0_DB_1534".Q AND ("Barcode462" > 0) AND "ปุ่มยืนยันหน้า Screen",
                           PV := 5,
                           CV => "Barcode462");
   "M462" := "IEC_Counter_0_DB_489".QU;
   "IEC_Counter_0_DB_1535".CTU(CU := "ยา 463" = 1,
                           R := "Stepper Motor ทำงาน สั่งconveyor เคลื่อที่ไปข้างหน้า" OR "ปุ่มClear",
                           PV := 1);
   "IEC_Counter_0_DB_490".CTUD(CU := ("Expected/Value_All".V = "Expected/Value_All".Expected_463) AND NOT "M463",
                           CD := "IEC_Counter_0_DB_1535".Q AND ("Barcode463" > 0) AND "ปุ่มยืนยันหน้า Screen",
                           PV := 5,
                           CV => "Barcode463");
   "M463" := "IEC_Counter_0_DB_490".QU;
   "IEC_Counter_0_DB_1536".CTU(CU := "ยา 464" = 1,
                           R := "Stepper Motor ทำงาน สั่งconveyor เคลื่อที่ไปข้างหน้า" OR "ปุ่มClear",
                           PV := 1);
   "IEC_Counter_0_DB_491".CTUD(CU := ("Expected/Value_All".V = "Expected/Value_All".Expected_464) AND NOT "M464",
                           CD := "IEC_Counter_0_DB_1536".Q AND ("Barcode464" > 0) AND "ปุ่มยืนยันหน้า Screen",
                           PV := 5,
                           CV => "Barcode464");
   "M464" := "IEC_Counter_0_DB_491".QU;
   "IEC_Counter_0_DB_1537".CTU(CU := "ยา 465" = 1,
                           R := "Stepper Motor ทำงาน สั่งconveyor เคลื่อที่ไปข้างหน้า" OR "ปุ่มClear",
                           PV := 1);
   "IEC_Counter_0_DB_492".CTUD(CU := ("Expected/Value_All".V = "Expected/Value_All".Expected_465) AND NOT "M465",
                           CD := "IEC_Counter_0_DB_1537".Q AND ("Barcode465" > 0) AND "ปุ่มยืนยันหน้า Screen",
                           PV := 5,
                           CV => "Barcode465");
   "M465" := "IEC_Counter_0_DB_492".QU;
   "IEC_Counter_0_DB_1538".CTU(CU := "ยา 466" = 1,
                           R := "Stepper Motor ทำงาน สั่งconveyor เคลื่อที่ไปข้างหน้า" OR "ปุ่มClear",
                           PV := 1);
   "IEC_Counter_0_DB_493".CTUD(CU := ("Expected/Value_All".V = "Expected/Value_All".Expected_466) AND NOT "M466",
                           CD := "IEC_Counter_0_DB_1538".Q AND ("Barcode466" > 0) AND "ปุ่มยืนยันหน้า Screen",
                           PV := 5,
                           CV => "Barcode466");
   "M466" := "IEC_Counter_0_DB_493".QU;
   "IEC_Counter_0_DB_1539".CTU(CU := "ยา 467" = 1,
                           R := "Stepper Motor ทำงาน สั่งconveyor เคลื่อที่ไปข้างหน้า" OR "ปุ่มClear",
                           PV := 1);
   "IEC_Counter_0_DB_494".CTUD(CU := ("Expected/Value_All".V = "Expected/Value_All".Expected_467) AND NOT "M467",
                           CD := "IEC_Counter_0_DB_1539".Q AND ("Barcode467" > 0) AND "ปุ่มยืนยันหน้า Screen",
                           PV := 5,
                           CV => "Barcode467");
   "M467" := "IEC_Counter_0_DB_494".QU;
   "IEC_Counter_0_DB_1540".CTU(CU := "ยา 468" = 1,
                           R := "Stepper Motor ทำงาน สั่งconveyor เคลื่อที่ไปข้างหน้า" OR "ปุ่มClear",
                           PV := 1);
   "IEC_Counter_0_DB_495".CTUD(CU := ("Expected/Value_All".V = "Expected/Value_All".Expected_468) AND NOT "M468",
                           CD := "IEC_Counter_0_DB_1540".Q AND ("Barcode468" > 0) AND "ปุ่มยืนยันหน้า Screen",
                           PV := 5,
                           CV => "Barcode468");
   "M468" := "IEC_Counter_0_DB_495".QU;
   "IEC_Counter_0_DB_1541".CTU(CU := "ยา 469" = 1,
                           R := "Stepper Motor ทำงาน สั่งconveyor เคลื่อที่ไปข้างหน้า" OR "ปุ่มClear",
                           PV := 1);
   "IEC_Counter_0_DB_496".CTUD(CU := ("Expected/Value_All".V = "Expected/Value_All".Expected_469) AND NOT "M469",
                           CD := "IEC_Counter_0_DB_1541".Q AND ("Barcode469" > 0) AND "ปุ่มยืนยันหน้า Screen",
                           PV := 5,
                           CV => "Barcode469");
   "M469" := "IEC_Counter_0_DB_496".QU;
   "IEC_Counter_0_DB_1542".CTU(CU := "ยา 470" = 1,
                           R := "Stepper Motor ทำงาน สั่งconveyor เคลื่อที่ไปข้างหน้า" OR "ปุ่มClear",
                           PV := 1);
   "IEC_Counter_0_DB_497".CTUD(CU := ("Expected/Value_All".V = "Expected/Value_All".Expected_470) AND NOT "M470",
                           CD := "IEC_Counter_0_DB_1542".Q AND ("Barcode470" > 0) AND "ปุ่มยืนยันหน้า Screen",
                           PV := 5,
                           CV => "Barcode470");
   "M470" := "IEC_Counter_0_DB_497".QU;
   "IEC_Counter_0_DB_1543".CTU(CU := "ยา 471" = 1,
                           R := "Stepper Motor ทำงาน สั่งconveyor เคลื่อที่ไปข้างหน้า" OR "ปุ่มClear",
                           PV := 1);
   "IEC_Counter_0_DB_498".CTUD(CU := ("Expected/Value_All".V = "Expected/Value_All".Expected_471) AND NOT "M471",
                           CD := "IEC_Counter_0_DB_1543".Q AND ("Barcode471" > 0) AND "ปุ่มยืนยันหน้า Screen",
                           PV := 5,
                           CV => "Barcode471");
   "M471" := "IEC_Counter_0_DB_498".QU;
   "IEC_Counter_0_DB_1544".CTU(CU := "ยา 472" = 1,
                           R := "Stepper Motor ทำงาน สั่งconveyor เคลื่อที่ไปข้างหน้า" OR "ปุ่มClear",
                           PV := 1);
   "IEC_Counter_0_DB_499".CTUD(CU := ("Expected/Value_All".V = "Expected/Value_All".Expected_472) AND NOT "M472",
                           CD := "IEC_Counter_0_DB_1544".Q AND ("Barcode472" > 0) AND "ปุ่มยืนยันหน้า Screen",
                           PV := 5,
                           CV => "Barcode472");
   "M472" := "IEC_Counter_0_DB_499".QU;
   "IEC_Counter_0_DB_1545".CTU(CU := "ยา 473" = 1,
                           R := "Stepper Motor ทำงาน สั่งconveyor เคลื่อที่ไปข้างหน้า" OR "ปุ่มClear",
                           PV := 1);
   "IEC_Counter_0_DB_500".CTUD(CU := ("Expected/Value_All".V = "Expected/Value_All".Expected_473) AND NOT "M473",
                           CD := "IEC_Counter_0_DB_1545".Q AND ("Barcode473" > 0) AND "ปุ่มยืนยันหน้า Screen",
                           PV := 5,
                           CV => "Barcode473");
   "M473" := "IEC_Counter_0_DB_500".QU;
   "IEC_Counter_0_DB_1546".CTU(CU := "ยา 474" = 1,
                           R := "Stepper Motor ทำงาน สั่งconveyor เคลื่อที่ไปข้างหน้า" OR "ปุ่มClear",
                           PV := 1);
   "IEC_Counter_0_DB_501".CTUD(CU := ("Expected/Value_All".V = "Expected/Value_All".Expected_474) AND NOT "M474",
                           CD := "IEC_Counter_0_DB_1546".Q AND ("Barcode474" > 0) AND "ปุ่มยืนยันหน้า Screen",
                           PV := 5,
                           CV => "Barcode474");
   "M474" := "IEC_Counter_0_DB_501".QU;
   "IEC_Counter_0_DB_1547".CTU(CU := "ยา 475" = 1,
                           R := "Stepper Motor ทำงาน สั่งconveyor เคลื่อที่ไปข้างหน้า" OR "ปุ่มClear",
                           PV := 1);
   "IEC_Counter_0_DB_502".CTUD(CU := ("Expected/Value_All".V = "Expected/Value_All".Expected_475) AND NOT "M475",
                           CD := "IEC_Counter_0_DB_1547".Q AND ("Barcode475" > 0) AND "ปุ่มยืนยันหน้า Screen",
                           PV := 5,
                           CV => "Barcode475");
   "M475" := "IEC_Counter_0_DB_502".QU;
   "IEC_Counter_0_DB_1548".CTU(CU := "ยา 476" = 1,
                           R := "Stepper Motor ทำงาน สั่งconveyor เคลื่อที่ไปข้างหน้า" OR "ปุ่มClear",
                           PV := 1);
   "IEC_Counter_0_DB_503".CTUD(CU := ("Expected/Value_All".V = "Expected/Value_All".Expected_476) AND NOT "M476",
                           CD := "IEC_Counter_0_DB_1548".Q AND ("Barcode476" > 0) AND "ปุ่มยืนยันหน้า Screen",
                           PV := 5,
                           CV => "Barcode476");
   "M476" := "IEC_Counter_0_DB_503".QU;
   "IEC_Counter_0_DB_1549".CTU(CU := "ยา 477" = 1,
                           R := "Stepper Motor ทำงาน สั่งconveyor เคลื่อที่ไปข้างหน้า" OR "ปุ่มClear",
                           PV := 1);
   "IEC_Counter_0_DB_504".CTUD(CU := ("Expected/Value_All".V = "Expected/Value_All".Expected_477) AND NOT "M477",
                           CD := "IEC_Counter_0_DB_1549".Q AND ("Barcode477" > 0) AND "ปุ่มยืนยันหน้า Screen",
                           PV := 5,
                           CV => "Barcode477");
   "M477" := "IEC_Counter_0_DB_504".QU;
   "IEC_Counter_0_DB_1550".CTU(CU := "ยา 478" = 1,
                           R := "Stepper Motor ทำงาน สั่งconveyor เคลื่อที่ไปข้างหน้า" OR "ปุ่มClear",
                           PV := 1);
   "IEC_Counter_0_DB_505".CTUD(CU := ("Expected/Value_All".V = "Expected/Value_All".Expected_478) AND NOT "M478",
                           CD := "IEC_Counter_0_DB_1550".Q AND ("Barcode478" > 0) AND "ปุ่มยืนยันหน้า Screen",
                           PV := 5,
                           CV => "Barcode478");
   "M478" := "IEC_Counter_0_DB_505".QU;
   "IEC_Counter_0_DB_1551".CTU(CU := "ยา 479" = 1,
                           R := "Stepper Motor ทำงาน สั่งconveyor เคลื่อที่ไปข้างหน้า" OR "ปุ่มClear",
                           PV := 1);
   "IEC_Counter_0_DB_506".CTUD(CU := ("Expected/Value_All".V = "Expected/Value_All".Expected_479) AND NOT "M479",
                           CD := "IEC_Counter_0_DB_1551".Q AND ("Barcode479" > 0) AND "ปุ่มยืนยันหน้า Screen",
                           PV := 5,
                           CV => "Barcode479");
   "M479" := "IEC_Counter_0_DB_506".QU;
   "IEC_Counter_0_DB_1552".CTU(CU := "ยา 480" = 1,
                           R := "Stepper Motor ทำงาน สั่งconveyor เคลื่อที่ไปข้างหน้า" OR "ปุ่มClear",
                           PV := 1);
   "IEC_Counter_0_DB_507".CTUD(CU := ("Expected/Value_All".V = "Expected/Value_All".Expected_480) AND NOT "M480",
                           CD := "IEC_Counter_0_DB_1552".Q AND ("Barcode480" > 0) AND "ปุ่มยืนยันหน้า Screen",
                           PV := 5,
                           CV => "Barcode480");
   "M480" := "IEC_Counter_0_DB_507".QU;
END_REGION

REGION Network 25
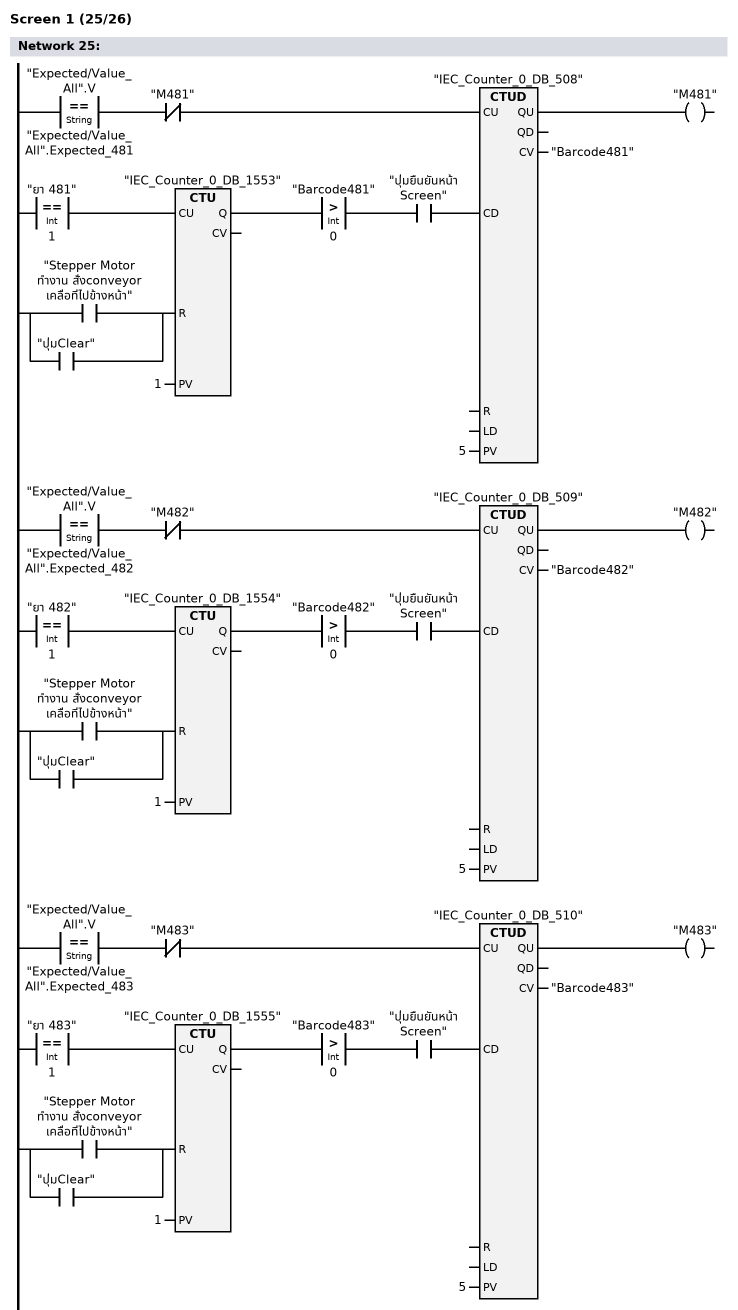
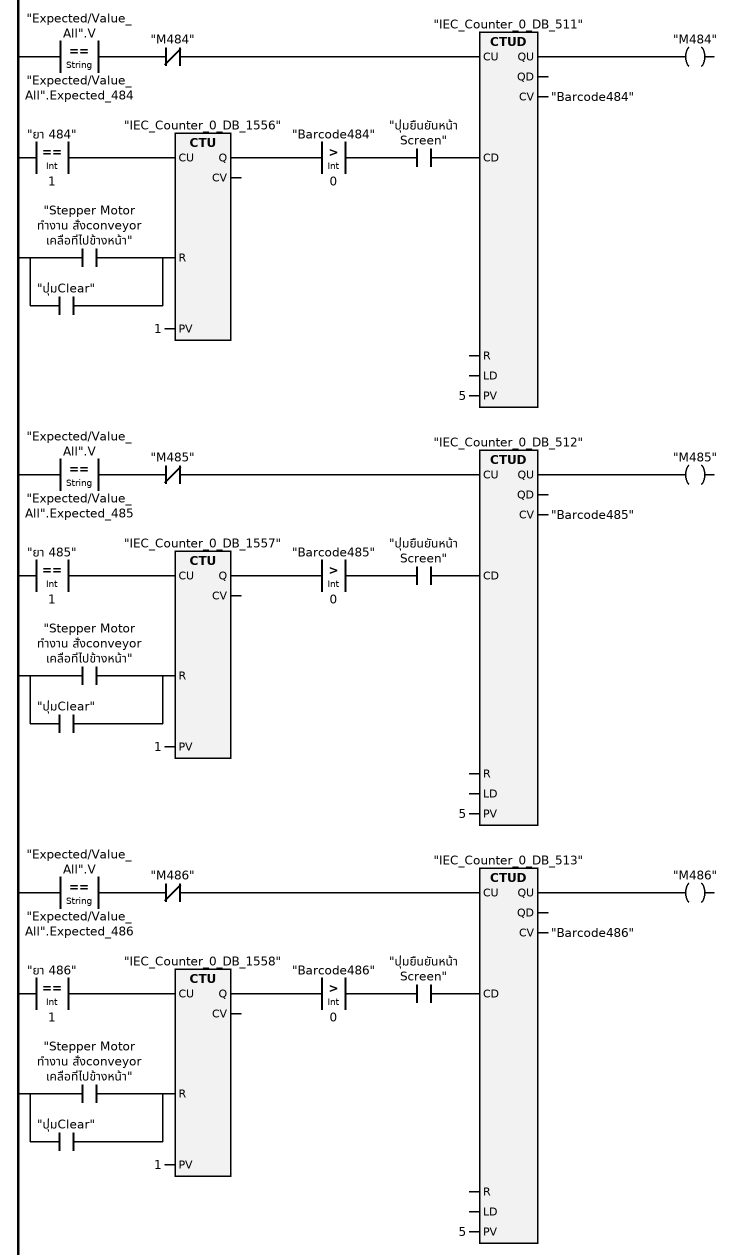
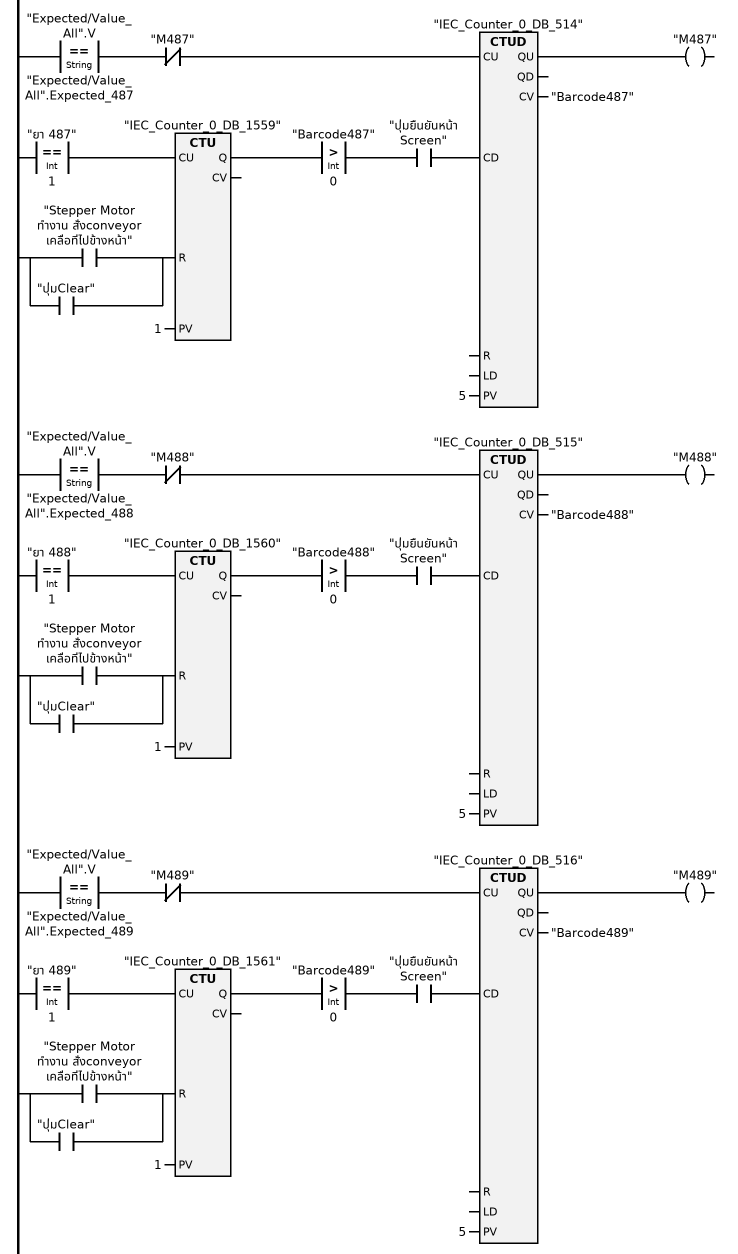
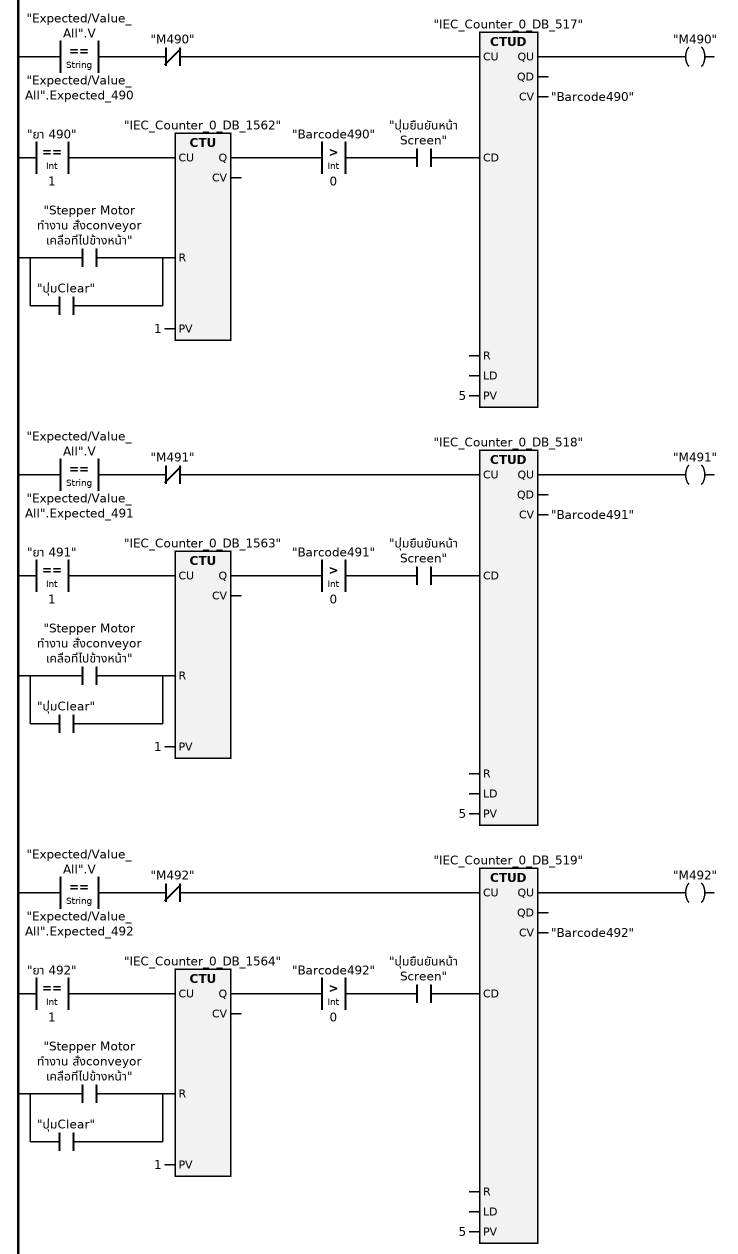
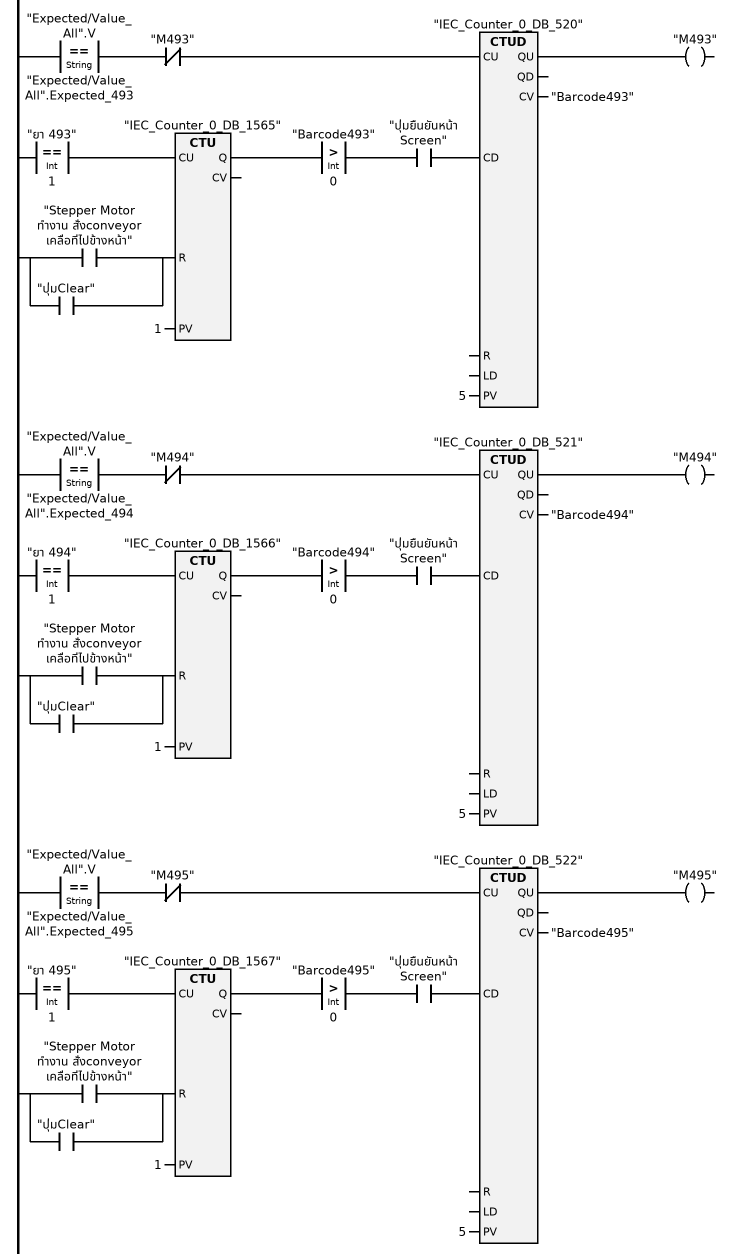
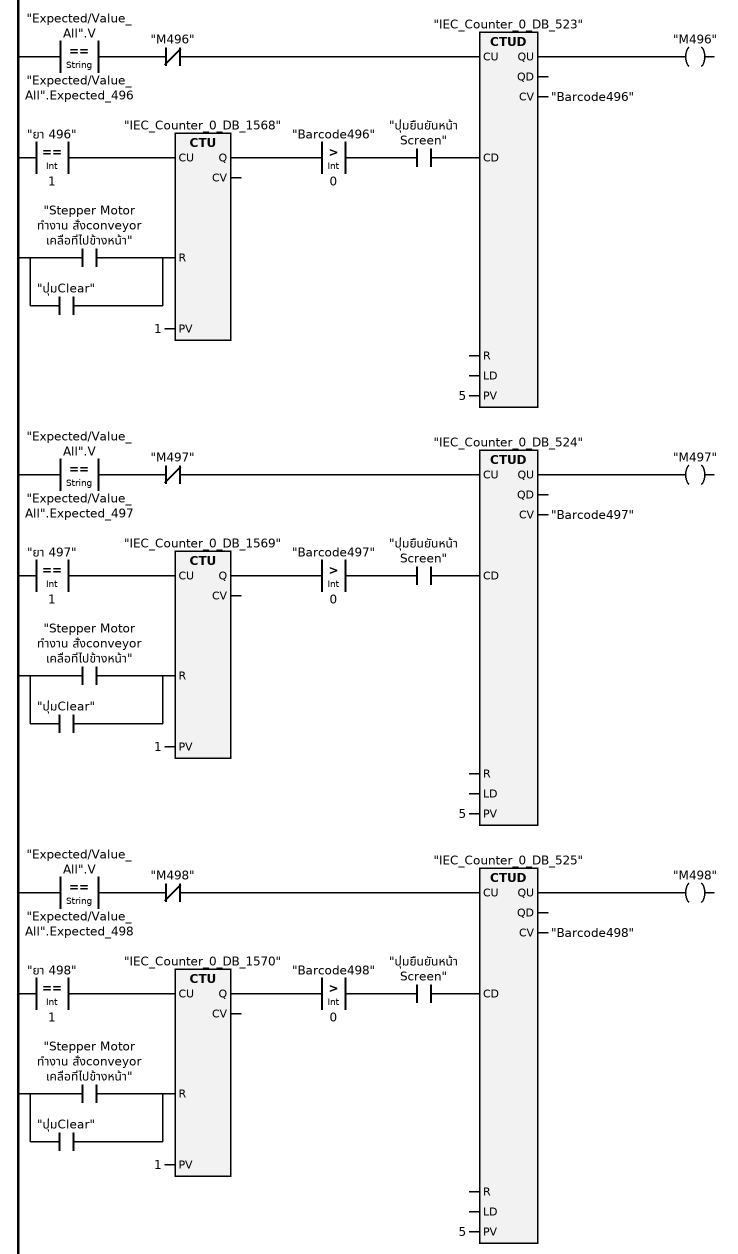
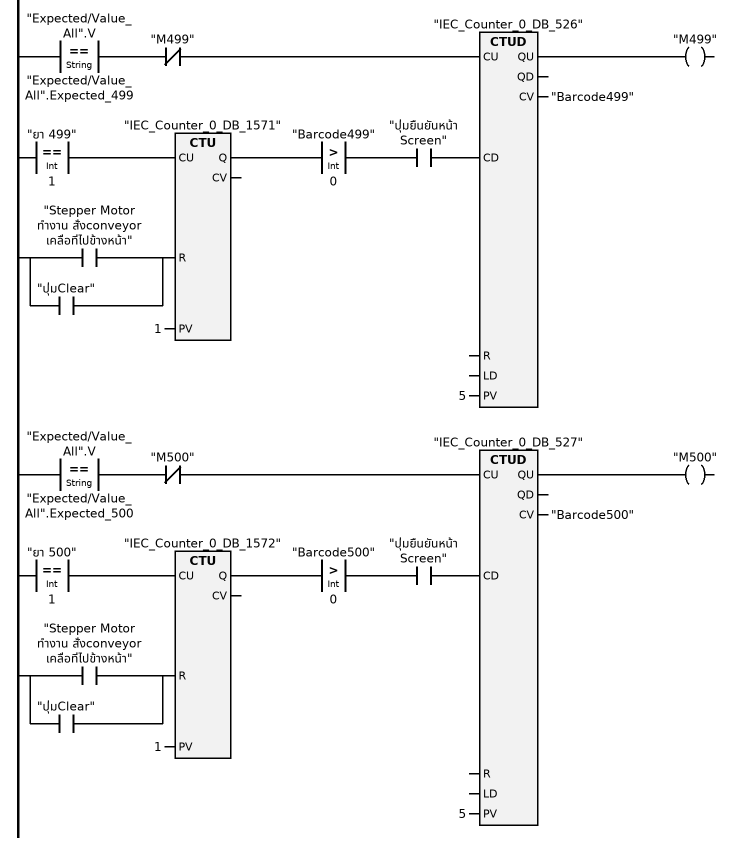
   "IEC_Counter_0_DB_1553".CTU(CU := "ยา 481" = 1,
                           R := "Stepper Motor ทำงาน สั่งconveyor เคลื่อที่ไปข้างหน้า" OR "ปุ่มClear",
                           PV := 1);
   "IEC_Counter_0_DB_508".CTUD(CU := ("Expected/Value_All".V = "Expected/Value_All".Expected_481) AND NOT "M481",
                           CD := "IEC_Counter_0_DB_1553".Q AND ("Barcode481" > 0) AND "ปุ่มยืนยันหน้า Screen",
                           PV := 5,
                           CV => "Barcode481");
   "M481" := "IEC_Counter_0_DB_508".QU;
   "IEC_Counter_0_DB_1554".CTU(CU := "ยา 482" = 1,
                           R := "Stepper Motor ทำงาน สั่งconveyor เคลื่อที่ไปข้างหน้า" OR "ปุ่มClear",
                           PV := 1);
   "IEC_Counter_0_DB_509".CTUD(CU := ("Expected/Value_All".V = "Expected/Value_All".Expected_482) AND NOT "M482",
                           CD := "IEC_Counter_0_DB_1554".Q AND ("Barcode482" > 0) AND "ปุ่มยืนยันหน้า Screen",
                           PV := 5,
                           CV => "Barcode482");
   "M482" := "IEC_Counter_0_DB_509".QU;
   "IEC_Counter_0_DB_1555".CTU(CU := "ยา 483" = 1,
                           R := "Stepper Motor ทำงาน สั่งconveyor เคลื่อที่ไปข้างหน้า" OR "ปุ่มClear",
                           PV := 1);
   "IEC_Counter_0_DB_510".CTUD(CU := ("Expected/Value_All".V = "Expected/Value_All".Expected_483) AND NOT "M483",
                           CD := "IEC_Counter_0_DB_1555".Q AND ("Barcode483" > 0) AND "ปุ่มยืนยันหน้า Screen",
                           PV := 5,
                           CV => "Barcode483");
   "M483" := "IEC_Counter_0_DB_510".QU;
   "IEC_Counter_0_DB_1556".CTU(CU := "ยา 484" = 1,
                           R := "Stepper Motor ทำงาน สั่งconveyor เคลื่อที่ไปข้างหน้า" OR "ปุ่มClear",
                           PV := 1);
   "IEC_Counter_0_DB_511".CTUD(CU := ("Expected/Value_All".V = "Expected/Value_All".Expected_484) AND NOT "M484",
                           CD := "IEC_Counter_0_DB_1556".Q AND ("Barcode484" > 0) AND "ปุ่มยืนยันหน้า Screen",
                           PV := 5,
                           CV => "Barcode484");
   "M484" := "IEC_Counter_0_DB_511".QU;
   "IEC_Counter_0_DB_1557".CTU(CU := "ยา 485" = 1,
                           R := "Stepper Motor ทำงาน สั่งconveyor เคลื่อที่ไปข้างหน้า" OR "ปุ่มClear",
                           PV := 1);
   "IEC_Counter_0_DB_512".CTUD(CU := ("Expected/Value_All".V = "Expected/Value_All".Expected_485) AND NOT "M485",
                           CD := "IEC_Counter_0_DB_1557".Q AND ("Barcode485" > 0) AND "ปุ่มยืนยันหน้า Screen",
                           PV := 5,
                           CV => "Barcode485");
   "M485" := "IEC_Counter_0_DB_512".QU;
   "IEC_Counter_0_DB_1558".CTU(CU := "ยา 486" = 1,
                           R := "Stepper Motor ทำงาน สั่งconveyor เคลื่อที่ไปข้างหน้า" OR "ปุ่มClear",
                           PV := 1);
   "IEC_Counter_0_DB_513".CTUD(CU := ("Expected/Value_All".V = "Expected/Value_All".Expected_486) AND NOT "M486",
                           CD := "IEC_Counter_0_DB_1558".Q AND ("Barcode486" > 0) AND "ปุ่มยืนยันหน้า Screen",
                           PV := 5,
                           CV => "Barcode486");
   "M486" := "IEC_Counter_0_DB_513".QU;
   "IEC_Counter_0_DB_1559".CTU(CU := "ยา 487" = 1,
                           R := "Stepper Motor ทำงาน สั่งconveyor เคลื่อที่ไปข้างหน้า" OR "ปุ่มClear",
                           PV := 1);
   "IEC_Counter_0_DB_514".CTUD(CU := ("Expected/Value_All".V = "Expected/Value_All".Expected_487) AND NOT "M487",
                           CD := "IEC_Counter_0_DB_1559".Q AND ("Barcode487" > 0) AND "ปุ่มยืนยันหน้า Screen",
                           PV := 5,
                           CV => "Barcode487");
   "M487" := "IEC_Counter_0_DB_514".QU;
   "IEC_Counter_0_DB_1560".CTU(CU := "ยา 488" = 1,
                           R := "Stepper Motor ทำงาน สั่งconveyor เคลื่อที่ไปข้างหน้า" OR "ปุ่มClear",
                           PV := 1);
   "IEC_Counter_0_DB_515".CTUD(CU := ("Expected/Value_All".V = "Expected/Value_All".Expected_488) AND NOT "M488",
                           CD := "IEC_Counter_0_DB_1560".Q AND ("Barcode488" > 0) AND "ปุ่มยืนยันหน้า Screen",
                           PV := 5,
                           CV => "Barcode488");
   "M488" := "IEC_Counter_0_DB_515".QU;
   "IEC_Counter_0_DB_1561".CTU(CU := "ยา 489" = 1,
                           R := "Stepper Motor ทำงาน สั่งconveyor เคลื่อที่ไปข้างหน้า" OR "ปุ่มClear",
                           PV := 1);
   "IEC_Counter_0_DB_516".CTUD(CU := ("Expected/Value_All".V = "Expected/Value_All".Expected_489) AND NOT "M489",
                           CD := "IEC_Counter_0_DB_1561".Q AND ("Barcode489" > 0) AND "ปุ่มยืนยันหน้า Screen",
                           PV := 5,
                           CV => "Barcode489");
   "M489" := "IEC_Counter_0_DB_516".QU;
   "IEC_Counter_0_DB_1562".CTU(CU := "ยา 490" = 1,
                           R := "Stepper Motor ทำงาน สั่งconveyor เคลื่อที่ไปข้างหน้า" OR "ปุ่มClear",
                           PV := 1);
   "IEC_Counter_0_DB_517".CTUD(CU := ("Expected/Value_All".V = "Expected/Value_All".Expected_490) AND NOT "M490",
                           CD := "IEC_Counter_0_DB_1562".Q AND ("Barcode490" > 0) AND "ปุ่มยืนยันหน้า Screen",
                           PV := 5,
                           CV => "Barcode490");
   "M490" := "IEC_Counter_0_DB_517".QU;
   "IEC_Counter_0_DB_1563".CTU(CU := "ยา 491" = 1,
                           R := "Stepper Motor ทำงาน สั่งconveyor เคลื่อที่ไปข้างหน้า" OR "ปุ่มClear",
                           PV := 1);
   "IEC_Counter_0_DB_518".CTUD(CU := ("Expected/Value_All".V = "Expected/Value_All".Expected_491) AND NOT "M491",
                           CD := "IEC_Counter_0_DB_1563".Q AND ("Barcode491" > 0) AND "ปุ่มยืนยันหน้า Screen",
                           PV := 5,
                           CV => "Barcode491");
   "M491" := "IEC_Counter_0_DB_518".QU;
   "IEC_Counter_0_DB_1564".CTU(CU := "ยา 492" = 1,
                           R := "Stepper Motor ทำงาน สั่งconveyor เคลื่อที่ไปข้างหน้า" OR "ปุ่มClear",
                           PV := 1);
   "IEC_Counter_0_DB_519".CTUD(CU := ("Expected/Value_All".V = "Expected/Value_All".Expected_492) AND NOT "M492",
                           CD := "IEC_Counter_0_DB_1564".Q AND ("Barcode492" > 0) AND "ปุ่มยืนยันหน้า Screen",
                           PV := 5,
                           CV => "Barcode492");
   "M492" := "IEC_Counter_0_DB_519".QU;
   "IEC_Counter_0_DB_1565".CTU(CU := "ยา 493" = 1,
                           R := "Stepper Motor ทำงาน สั่งconveyor เคลื่อที่ไปข้างหน้า" OR "ปุ่มClear",
                           PV := 1);
   "IEC_Counter_0_DB_520".CTUD(CU := ("Expected/Value_All".V = "Expected/Value_All".Expected_493) AND NOT "M493",
                           CD := "IEC_Counter_0_DB_1565".Q AND ("Barcode493" > 0) AND "ปุ่มยืนยันหน้า Screen",
                           PV := 5,
                           CV => "Barcode493");
   "M493" := "IEC_Counter_0_DB_520".QU;
   "IEC_Counter_0_DB_1566".CTU(CU := "ยา 494" = 1,
                           R := "Stepper Motor ทำงาน สั่งconveyor เคลื่อที่ไปข้างหน้า" OR "ปุ่มClear",
                           PV := 1);
   "IEC_Counter_0_DB_521".CTUD(CU := ("Expected/Value_All".V = "Expected/Value_All".Expected_494) AND NOT "M494",
                           CD := "IEC_Counter_0_DB_1566".Q AND ("Barcode494" > 0) AND "ปุ่มยืนยันหน้า Screen",
                           PV := 5,
                           CV => "Barcode494");
   "M494" := "IEC_Counter_0_DB_521".QU;
   "IEC_Counter_0_DB_1567".CTU(CU := "ยา 495" = 1,
                           R := "Stepper Motor ทำงาน สั่งconveyor เคลื่อที่ไปข้างหน้า" OR "ปุ่มClear",
                           PV := 1);
   "IEC_Counter_0_DB_522".CTUD(CU := ("Expected/Value_All".V = "Expected/Value_All".Expected_495) AND NOT "M495",
                           CD := "IEC_Counter_0_DB_1567".Q AND ("Barcode495" > 0) AND "ปุ่มยืนยันหน้า Screen",
                           PV := 5,
                           CV => "Barcode495");
   "M495" := "IEC_Counter_0_DB_522".QU;
   "IEC_Counter_0_DB_1568".CTU(CU := "ยา 496" = 1,
                           R := "Stepper Motor ทำงาน สั่งconveyor เคลื่อที่ไปข้างหน้า" OR "ปุ่มClear",
                           PV := 1);
   "IEC_Counter_0_DB_523".CTUD(CU := ("Expected/Value_All".V = "Expected/Value_All".Expected_496) AND NOT "M496",
                           CD := "IEC_Counter_0_DB_1568".Q AND ("Barcode496" > 0) AND "ปุ่มยืนยันหน้า Screen",
                           PV := 5,
                           CV => "Barcode496");
   "M496" := "IEC_Counter_0_DB_523".QU;
   "IEC_Counter_0_DB_1569".CTU(CU := "ยา 497" = 1,
                           R := "Stepper Motor ทำงาน สั่งconveyor เคลื่อที่ไปข้างหน้า" OR "ปุ่มClear",
                           PV := 1);
   "IEC_Counter_0_DB_524".CTUD(CU := ("Expected/Value_All".V = "Expected/Value_All".Expected_497) AND NOT "M497",
                           CD := "IEC_Counter_0_DB_1569".Q AND ("Barcode497" > 0) AND "ปุ่มยืนยันหน้า Screen",
                           PV := 5,
                           CV => "Barcode497");
   "M497" := "IEC_Counter_0_DB_524".QU;
   "IEC_Counter_0_DB_1570".CTU(CU := "ยา 498" = 1,
                           R := "Stepper Motor ทำงาน สั่งconveyor เคลื่อที่ไปข้างหน้า" OR "ปุ่มClear",
                           PV := 1);
   "IEC_Counter_0_DB_525".CTUD(CU := ("Expected/Value_All".V = "Expected/Value_All".Expected_498) AND NOT "M498",
                           CD := "IEC_Counter_0_DB_1570".Q AND ("Barcode498" > 0) AND "ปุ่มยืนยันหน้า Screen",
                           PV := 5,
                           CV => "Barcode498");
   "M498" := "IEC_Counter_0_DB_525".QU;
   "IEC_Counter_0_DB_1571".CTU(CU := "ยา 499" = 1,
                           R := "Stepper Motor ทำงาน สั่งconveyor เคลื่อที่ไปข้างหน้า" OR "ปุ่มClear",
                           PV := 1);
   "IEC_Counter_0_DB_526".CTUD(CU := ("Expected/Value_All".V = "Expected/Value_All".Expected_499) AND NOT "M499",
                           CD := "IEC_Counter_0_DB_1571".Q AND ("Barcode499" > 0) AND "ปุ่มยืนยันหน้า Screen",
                           PV := 5,
                           CV => "Barcode499");
   "M499" := "IEC_Counter_0_DB_526".QU;
   "IEC_Counter_0_DB_1572".CTU(CU := "ยา 500" = 1,
                           R := "Stepper Motor ทำงาน สั่งconveyor เคลื่อที่ไปข้างหน้า" OR "ปุ่มClear",
                           PV := 1);
   "IEC_Counter_0_DB_527".CTUD(CU := ("Expected/Value_All".V = "Expected/Value_All".Expected_500) AND NOT "M500",
                           CD := "IEC_Counter_0_DB_1572".Q AND ("Barcode500" > 0) AND "ปุ่มยืนยันหน้า Screen",
                           PV := 5,
                           CV => "Barcode500");
   "M500" := "IEC_Counter_0_DB_527".QU;
END_REGION

REGION Network 26
